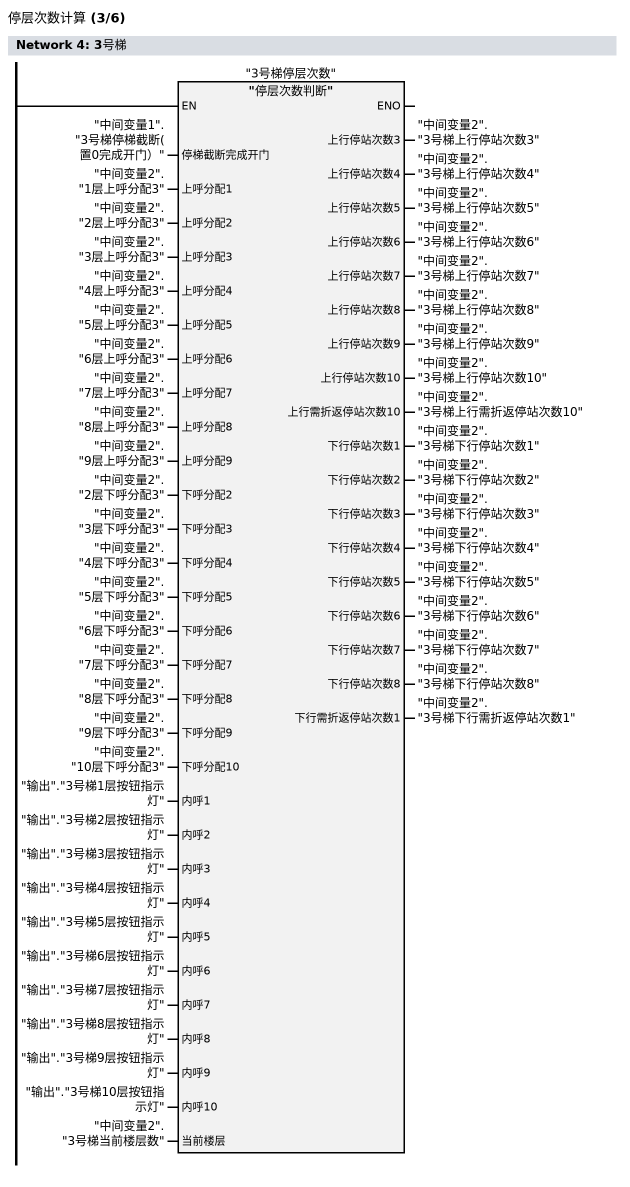
   RUNG wire#powerrail
      "3号梯停层次数"(停梯截断完成开门 := "中间变量1"."3号梯停梯截断(置0完成开门）", 上呼分配1 := "中间变量2"."1层上呼分配3", 上呼分配2 := "中间变量2"."2层上呼分配3", 上呼分配3 := "中间变量2"."3层上呼分配3", 上呼分配4 := "中间变量2"."4层上呼分配3", 上呼分配5 := "中间变量2"."5层上呼分配3", 上呼分配6 := "中间变量2"."6层上呼分配3", 上呼分配7 := "中间变量2"."7层上呼分配3", 上呼分配8 := "中间变量2"."8层上呼分配3", 上呼分配9 := "中间变量2"."9层上呼分配3", 下呼分配2 := "中间变量2"."2层下呼分配3", 下呼分配3 := "中间变量2"."3层下呼分配3", 下呼分配4 := "中间变量2"."4层下呼分配3", 下呼分配5 := "中间变量2"."5层下呼分配3", 下呼分配6 := "中间变量2"."6层下呼分配3", 下呼分配7 := "中间变量2"."7层下呼分配3", 下呼分配8 := "中间变量2"."8层下呼分配3", 下呼分配9 := "中间变量2"."9层下呼分配3", 下呼分配10 := "中间变量2"."10层下呼分配3", 内呼1 := "输出"."3号梯1层按钮指示灯", 内呼2 := "输出"."3号梯2层按钮指示灯", 内呼3 := "输出"."3号梯3层按钮指示灯", 内呼4 := "输出"."3号梯4层按钮指示灯", 内呼5 := "输出"."3号梯5层按钮指示灯", 内呼6 := "输出"."3号梯6层按钮指示灯", 内呼7 := "输出"."3号梯7层按钮指示灯", 内呼8 := "输出"."3号梯8层按钮指示灯", 内呼9 := "输出"."3号梯9层按钮指示灯", 内呼10 := "输出"."3号梯10层按钮指示灯", 当前楼层 := "中间变量2"."3号梯当前楼层数", 上行停站次数3 => "中间变量2"."3号梯上行停站次数3", 上行停站次数4 => "中间变量2"."3号梯上行停站次数4", 上行停站次数5 => "中间变量2"."3号梯上行停站次数5", 上行停站次数6 => "中间变量2"."3号梯上行停站次数6", 上行停站次数7 => "中间变量2"."3号梯上行停站次数7", 上行停站次数8 => "中间变量2"."3号梯上行停站次数8", 上行停站次数9 => "中间变量2"."3号梯上行停站次数9", 上行停站次数10 => "中间变量2"."3号梯上行停站次数10", 上行需折返停站次数10 => "中间变量2"."3号梯上行需折返停站次数10", 下行停站次数1 => "中间变量2"."3号梯下行停站次数1", 下行停站次数2 => "中间变量2"."3号梯下行停站次数2", 下行停站次数3 => "中间变量2"."3号梯下行停站次数3", 下行停站次数4 => "中间变量2"."3号梯下行停站次数4", 下行停站次数5 => "中间变量2"."3号梯下行停站次数5", 下行停站次数6 => "中间变量2"."3号梯下行停站次数6", 下行停站次数7 => "中间变量2"."3号梯下行停站次数7", 下行停站次数8 => "中间变量2"."3号梯下行停站次数8", 下行需折返停站次数1 => "中间变量2"."3号梯下行需折返停站次数1")
   END_RUNG
   // the same network as SCL:
   "3号梯停层次数"(停梯截断完成开门 := "中间变量1"."3号梯停梯截断(置0完成开门）",   // "停层次数判断"
             上呼分配1 := "中间变量2"."1层上呼分配3",
             上呼分配2 := "中间变量2"."2层上呼分配3",
             上呼分配3 := "中间变量2"."3层上呼分配3",
             上呼分配4 := "中间变量2"."4层上呼分配3",
             上呼分配5 := "中间变量2"."5层上呼分配3",
             上呼分配6 := "中间变量2"."6层上呼分配3",
             上呼分配7 := "中间变量2"."7层上呼分配3",
             上呼分配8 := "中间变量2"."8层上呼分配3",
             上呼分配9 := "中间变量2"."9层上呼分配3",
             下呼分配2 := "中间变量2"."2层下呼分配3",
             下呼分配3 := "中间变量2"."3层下呼分配3",
             下呼分配4 := "中间变量2"."4层下呼分配3",
             下呼分配5 := "中间变量2"."5层下呼分配3",
             下呼分配6 := "中间变量2"."6层下呼分配3",
             下呼分配7 := "中间变量2"."7层下呼分配3",
             下呼分配8 := "中间变量2"."8层下呼分配3",
             下呼分配9 := "中间变量2"."9层下呼分配3",
             下呼分配10 := "中间变量2"."10层下呼分配3",
             内呼1 := "输出"."3号梯1层按钮指示灯",
             内呼2 := "输出"."3号梯2层按钮指示灯",
             内呼3 := "输出"."3号梯3层按钮指示灯",
             内呼4 := "输出"."3号梯4层按钮指示灯",
             内呼5 := "输出"."3号梯5层按钮指示灯",
             内呼6 := "输出"."3号梯6层按钮指示灯",
             内呼7 := "输出"."3号梯7层按钮指示灯",
             内呼8 := "输出"."3号梯8层按钮指示灯",
             内呼9 := "输出"."3号梯9层按钮指示灯",
             内呼10 := "输出"."3号梯10层按钮指示灯",
             当前楼层 := "中间变量2"."3号梯当前楼层数",
             上行停站次数3 => "中间变量2"."3号梯上行停站次数3",
             上行停站次数4 => "中间变量2"."3号梯上行停站次数4",
             上行停站次数5 => "中间变量2"."3号梯上行停站次数5",
             上行停站次数6 => "中间变量2"."3号梯上行停站次数6",
             上行停站次数7 => "中间变量2"."3号梯上行停站次数7",
             上行停站次数8 => "中间变量2"."3号梯上行停站次数8",
             上行停站次数9 => "中间变量2"."3号梯上行停站次数9",
             上行停站次数10 => "中间变量2"."3号梯上行停站次数10",
             上行需折返停站次数10 => "中间变量2"."3号梯上行需折返停站次数10",
             下行停站次数1 => "中间变量2"."3号梯下行停站次数1",
             下行停站次数2 => "中间变量2"."3号梯下行停站次数2",
             下行停站次数3 => "中间变量2"."3号梯下行停站次数3",
             下行停站次数4 => "中间变量2"."3号梯下行停站次数4",
             下行停站次数5 => "中间变量2"."3号梯下行停站次数5",
             下行停站次数6 => "中间变量2"."3号梯下行停站次数6",
             下行停站次数7 => "中间变量2"."3号梯下行停站次数7",
             下行停站次数8 => "中间变量2"."3号梯下行停站次数8",
             下行需折返停站次数1 => "中间变量2"."3号梯下行需折返停站次数1");
END_REGION

REGION Network 5: 4号梯
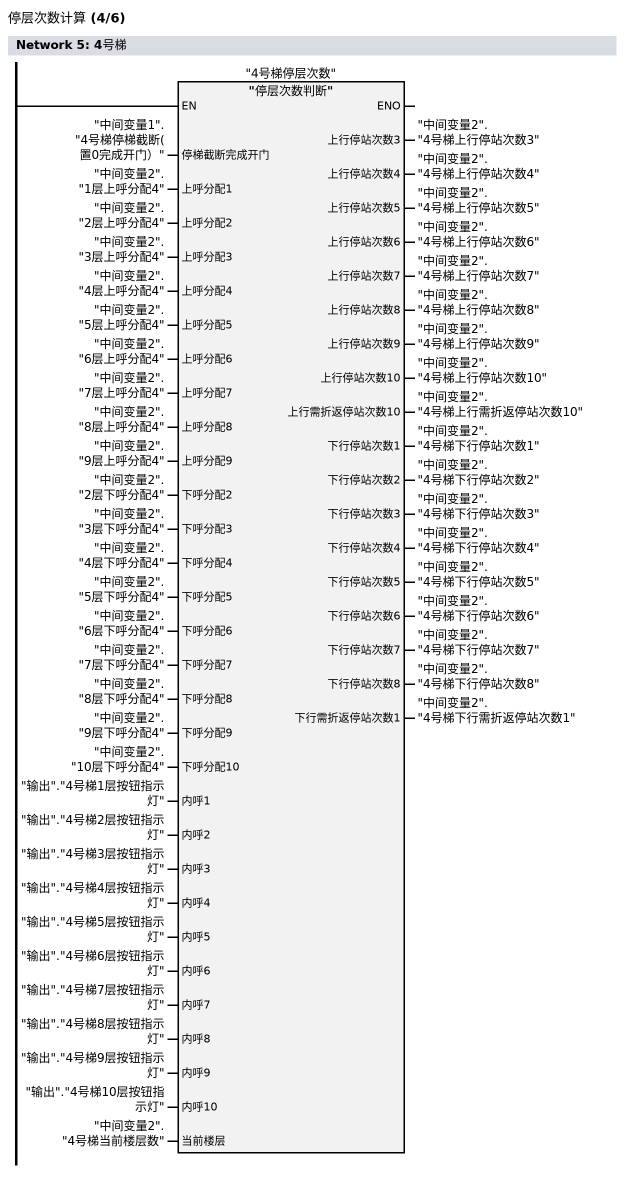
   RUNG wire#powerrail
      "4号梯停层次数"(停梯截断完成开门 := "中间变量1"."4号梯停梯截断(置0完成开门）", 上呼分配1 := "中间变量2"."1层上呼分配4", 上呼分配2 := "中间变量2"."2层上呼分配4", 上呼分配3 := "中间变量2"."3层上呼分配4", 上呼分配4 := "中间变量2"."4层上呼分配4", 上呼分配5 := "中间变量2"."5层上呼分配4", 上呼分配6 := "中间变量2"."6层上呼分配4", 上呼分配7 := "中间变量2"."7层上呼分配4", 上呼分配8 := "中间变量2"."8层上呼分配4", 上呼分配9 := "中间变量2"."9层上呼分配4", 下呼分配2 := "中间变量2"."2层下呼分配4", 下呼分配3 := "中间变量2"."3层下呼分配4", 下呼分配4 := "中间变量2"."4层下呼分配4", 下呼分配5 := "中间变量2"."5层下呼分配4", 下呼分配6 := "中间变量2"."6层下呼分配4", 下呼分配7 := "中间变量2"."7层下呼分配4", 下呼分配8 := "中间变量2"."8层下呼分配4", 下呼分配9 := "中间变量2"."9层下呼分配4", 下呼分配10 := "中间变量2"."10层下呼分配4", 内呼1 := "输出"."4号梯1层按钮指示灯", 内呼2 := "输出"."4号梯2层按钮指示灯", 内呼3 := "输出"."4号梯3层按钮指示灯", 内呼4 := "输出"."4号梯4层按钮指示灯", 内呼5 := "输出"."4号梯5层按钮指示灯", 内呼6 := "输出"."4号梯6层按钮指示灯", 内呼7 := "输出"."4号梯7层按钮指示灯", 内呼8 := "输出"."4号梯8层按钮指示灯", 内呼9 := "输出"."4号梯9层按钮指示灯", 内呼10 := "输出"."4号梯10层按钮指示灯", 当前楼层 := "中间变量2"."4号梯当前楼层数", 上行停站次数3 => "中间变量2"."4号梯上行停站次数3", 上行停站次数4 => "中间变量2"."4号梯上行停站次数4", 上行停站次数5 => "中间变量2"."4号梯上行停站次数5", 上行停站次数6 => "中间变量2"."4号梯上行停站次数6", 上行停站次数7 => "中间变量2"."4号梯上行停站次数7", 上行停站次数8 => "中间变量2"."4号梯上行停站次数8", 上行停站次数9 => "中间变量2"."4号梯上行停站次数9", 上行停站次数10 => "中间变量2"."4号梯上行停站次数10", 上行需折返停站次数10 => "中间变量2"."4号梯上行需折返停站次数10", 下行停站次数1 => "中间变量2"."4号梯下行停站次数1", 下行停站次数2 => "中间变量2"."4号梯下行停站次数2", 下行停站次数3 => "中间变量2"."4号梯下行停站次数3", 下行停站次数4 => "中间变量2"."4号梯下行停站次数4", 下行停站次数5 => "中间变量2"."4号梯下行停站次数5", 下行停站次数6 => "中间变量2"."4号梯下行停站次数6", 下行停站次数7 => "中间变量2"."4号梯下行停站次数7", 下行停站次数8 => "中间变量2"."4号梯下行停站次数8", 下行需折返停站次数1 => "中间变量2"."4号梯下行需折返停站次数1")
   END_RUNG
   // the same network as SCL:
   "4号梯停层次数"(停梯截断完成开门 := "中间变量1"."4号梯停梯截断(置0完成开门）",   // "停层次数判断"
             上呼分配1 := "中间变量2"."1层上呼分配4",
             上呼分配2 := "中间变量2"."2层上呼分配4",
             上呼分配3 := "中间变量2"."3层上呼分配4",
             上呼分配4 := "中间变量2"."4层上呼分配4",
             上呼分配5 := "中间变量2"."5层上呼分配4",
             上呼分配6 := "中间变量2"."6层上呼分配4",
             上呼分配7 := "中间变量2"."7层上呼分配4",
             上呼分配8 := "中间变量2"."8层上呼分配4",
             上呼分配9 := "中间变量2"."9层上呼分配4",
             下呼分配2 := "中间变量2"."2层下呼分配4",
             下呼分配3 := "中间变量2"."3层下呼分配4",
             下呼分配4 := "中间变量2"."4层下呼分配4",
             下呼分配5 := "中间变量2"."5层下呼分配4",
             下呼分配6 := "中间变量2"."6层下呼分配4",
             下呼分配7 := "中间变量2"."7层下呼分配4",
             下呼分配8 := "中间变量2"."8层下呼分配4",
             下呼分配9 := "中间变量2"."9层下呼分配4",
             下呼分配10 := "中间变量2"."10层下呼分配4",
             内呼1 := "输出"."4号梯1层按钮指示灯",
             内呼2 := "输出"."4号梯2层按钮指示灯",
             内呼3 := "输出"."4号梯3层按钮指示灯",
             内呼4 := "输出"."4号梯4层按钮指示灯",
             内呼5 := "输出"."4号梯5层按钮指示灯",
             内呼6 := "输出"."4号梯6层按钮指示灯",
             内呼7 := "输出"."4号梯7层按钮指示灯",
             内呼8 := "输出"."4号梯8层按钮指示灯",
             内呼9 := "输出"."4号梯9层按钮指示灯",
             内呼10 := "输出"."4号梯10层按钮指示灯",
             当前楼层 := "中间变量2"."4号梯当前楼层数",
             上行停站次数3 => "中间变量2"."4号梯上行停站次数3",
             上行停站次数4 => "中间变量2"."4号梯上行停站次数4",
             上行停站次数5 => "中间变量2"."4号梯上行停站次数5",
             上行停站次数6 => "中间变量2"."4号梯上行停站次数6",
             上行停站次数7 => "中间变量2"."4号梯上行停站次数7",
             上行停站次数8 => "中间变量2"."4号梯上行停站次数8",
             上行停站次数9 => "中间变量2"."4号梯上行停站次数9",
             上行停站次数10 => "中间变量2"."4号梯上行停站次数10",
             上行需折返停站次数10 => "中间变量2"."4号梯上行需折返停站次数10",
             下行停站次数1 => "中间变量2"."4号梯下行停站次数1",
             下行停站次数2 => "中间变量2"."4号梯下行停站次数2",
             下行停站次数3 => "中间变量2"."4号梯下行停站次数3",
             下行停站次数4 => "中间变量2"."4号梯下行停站次数4",
             下行停站次数5 => "中间变量2"."4号梯下行停站次数5",
             下行停站次数6 => "中间变量2"."4号梯下行停站次数6",
             下行停站次数7 => "中间变量2"."4号梯下行停站次数7",
             下行停站次数8 => "中间变量2"."4号梯下行停站次数8",
             下行需折返停站次数1 => "中间变量2"."4号梯下行需折返停站次数1");
END_REGION

REGION Network 6: 5号梯
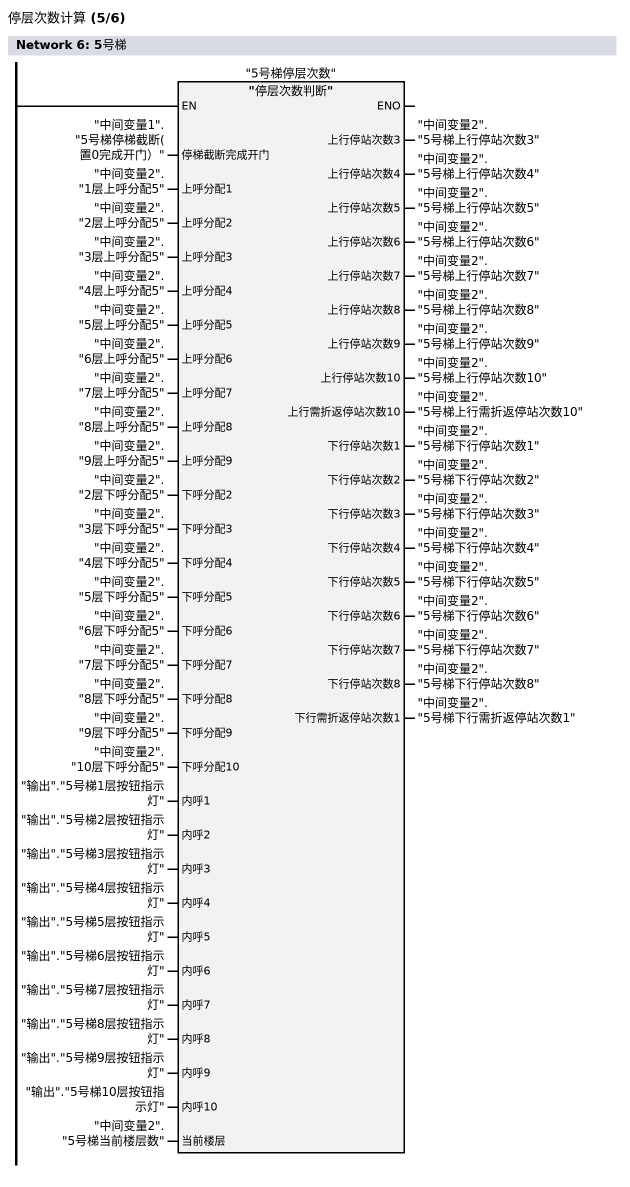
   RUNG wire#powerrail
      "5号梯停层次数"(停梯截断完成开门 := "中间变量1"."5号梯停梯截断(置0完成开门）", 上呼分配1 := "中间变量2"."1层上呼分配5", 上呼分配2 := "中间变量2"."2层上呼分配5", 上呼分配3 := "中间变量2"."3层上呼分配5", 上呼分配4 := "中间变量2"."4层上呼分配5", 上呼分配5 := "中间变量2"."5层上呼分配5", 上呼分配6 := "中间变量2"."6层上呼分配5", 上呼分配7 := "中间变量2"."7层上呼分配5", 上呼分配8 := "中间变量2"."8层上呼分配5", 上呼分配9 := "中间变量2"."9层上呼分配5", 下呼分配2 := "中间变量2"."2层下呼分配5", 下呼分配3 := "中间变量2"."3层下呼分配5", 下呼分配4 := "中间变量2"."4层下呼分配5", 下呼分配5 := "中间变量2"."5层下呼分配5", 下呼分配6 := "中间变量2"."6层下呼分配5", 下呼分配7 := "中间变量2"."7层下呼分配5", 下呼分配8 := "中间变量2"."8层下呼分配5", 下呼分配9 := "中间变量2"."9层下呼分配5", 下呼分配10 := "中间变量2"."10层下呼分配5", 内呼1 := "输出"."5号梯1层按钮指示灯", 内呼2 := "输出"."5号梯2层按钮指示灯", 内呼3 := "输出"."5号梯3层按钮指示灯", 内呼4 := "输出"."5号梯4层按钮指示灯", 内呼5 := "输出"."5号梯5层按钮指示灯", 内呼6 := "输出"."5号梯6层按钮指示灯", 内呼7 := "输出"."5号梯7层按钮指示灯", 内呼8 := "输出"."5号梯8层按钮指示灯", 内呼9 := "输出"."5号梯9层按钮指示灯", 内呼10 := "输出"."5号梯10层按钮指示灯", 当前楼层 := "中间变量2"."5号梯当前楼层数", 上行停站次数3 => "中间变量2"."5号梯上行停站次数3", 上行停站次数4 => "中间变量2"."5号梯上行停站次数4", 上行停站次数5 => "中间变量2"."5号梯上行停站次数5", 上行停站次数6 => "中间变量2"."5号梯上行停站次数6", 上行停站次数7 => "中间变量2"."5号梯上行停站次数7", 上行停站次数8 => "中间变量2"."5号梯上行停站次数8", 上行停站次数9 => "中间变量2"."5号梯上行停站次数9", 上行停站次数10 => "中间变量2"."5号梯上行停站次数10", 上行需折返停站次数10 => "中间变量2"."5号梯上行需折返停站次数10", 下行停站次数1 => "中间变量2"."5号梯下行停站次数1", 下行停站次数2 => "中间变量2"."5号梯下行停站次数2", 下行停站次数3 => "中间变量2"."5号梯下行停站次数3", 下行停站次数4 => "中间变量2"."5号梯下行停站次数4", 下行停站次数5 => "中间变量2"."5号梯下行停站次数5", 下行停站次数6 => "中间变量2"."5号梯下行停站次数6", 下行停站次数7 => "中间变量2"."5号梯下行停站次数7", 下行停站次数8 => "中间变量2"."5号梯下行停站次数8", 下行需折返停站次数1 => "中间变量2"."5号梯下行需折返停站次数1")
   END_RUNG
   // the same network as SCL:
   "5号梯停层次数"(停梯截断完成开门 := "中间变量1"."5号梯停梯截断(置0完成开门）",   // "停层次数判断"
             上呼分配1 := "中间变量2"."1层上呼分配5",
             上呼分配2 := "中间变量2"."2层上呼分配5",
             上呼分配3 := "中间变量2"."3层上呼分配5",
             上呼分配4 := "中间变量2"."4层上呼分配5",
             上呼分配5 := "中间变量2"."5层上呼分配5",
             上呼分配6 := "中间变量2"."6层上呼分配5",
             上呼分配7 := "中间变量2"."7层上呼分配5",
             上呼分配8 := "中间变量2"."8层上呼分配5",
             上呼分配9 := "中间变量2"."9层上呼分配5",
             下呼分配2 := "中间变量2"."2层下呼分配5",
             下呼分配3 := "中间变量2"."3层下呼分配5",
             下呼分配4 := "中间变量2"."4层下呼分配5",
             下呼分配5 := "中间变量2"."5层下呼分配5",
             下呼分配6 := "中间变量2"."6层下呼分配5",
             下呼分配7 := "中间变量2"."7层下呼分配5",
             下呼分配8 := "中间变量2"."8层下呼分配5",
             下呼分配9 := "中间变量2"."9层下呼分配5",
             下呼分配10 := "中间变量2"."10层下呼分配5",
             内呼1 := "输出"."5号梯1层按钮指示灯",
             内呼2 := "输出"."5号梯2层按钮指示灯",
             内呼3 := "输出"."5号梯3层按钮指示灯",
             内呼4 := "输出"."5号梯4层按钮指示灯",
             内呼5 := "输出"."5号梯5层按钮指示灯",
             内呼6 := "输出"."5号梯6层按钮指示灯",
             内呼7 := "输出"."5号梯7层按钮指示灯",
             内呼8 := "输出"."5号梯8层按钮指示灯",
             内呼9 := "输出"."5号梯9层按钮指示灯",
             内呼10 := "输出"."5号梯10层按钮指示灯",
             当前楼层 := "中间变量2"."5号梯当前楼层数",
             上行停站次数3 => "中间变量2"."5号梯上行停站次数3",
             上行停站次数4 => "中间变量2"."5号梯上行停站次数4",
             上行停站次数5 => "中间变量2"."5号梯上行停站次数5",
             上行停站次数6 => "中间变量2"."5号梯上行停站次数6",
             上行停站次数7 => "中间变量2"."5号梯上行停站次数7",
             上行停站次数8 => "中间变量2"."5号梯上行停站次数8",
             上行停站次数9 => "中间变量2"."5号梯上行停站次数9",
             上行停站次数10 => "中间变量2"."5号梯上行停站次数10",
             上行需折返停站次数10 => "中间变量2"."5号梯上行需折返停站次数10",
             下行停站次数1 => "中间变量2"."5号梯下行停站次数1",
             下行停站次数2 => "中间变量2"."5号梯下行停站次数2",
             下行停站次数3 => "中间变量2"."5号梯下行停站次数3",
             下行停站次数4 => "中间变量2"."5号梯下行停站次数4",
             下行停站次数5 => "中间变量2"."5号梯下行停站次数5",
             下行停站次数6 => "中间变量2"."5号梯下行停站次数6",
             下行停站次数7 => "中间变量2"."5号梯下行停站次数7",
             下行停站次数8 => "中间变量2"."5号梯下行停站次数8",
             下行需折返停站次数1 => "中间变量2"."5号梯下行需折返停站次数1");
END_REGION

REGION Network 7: 6号梯
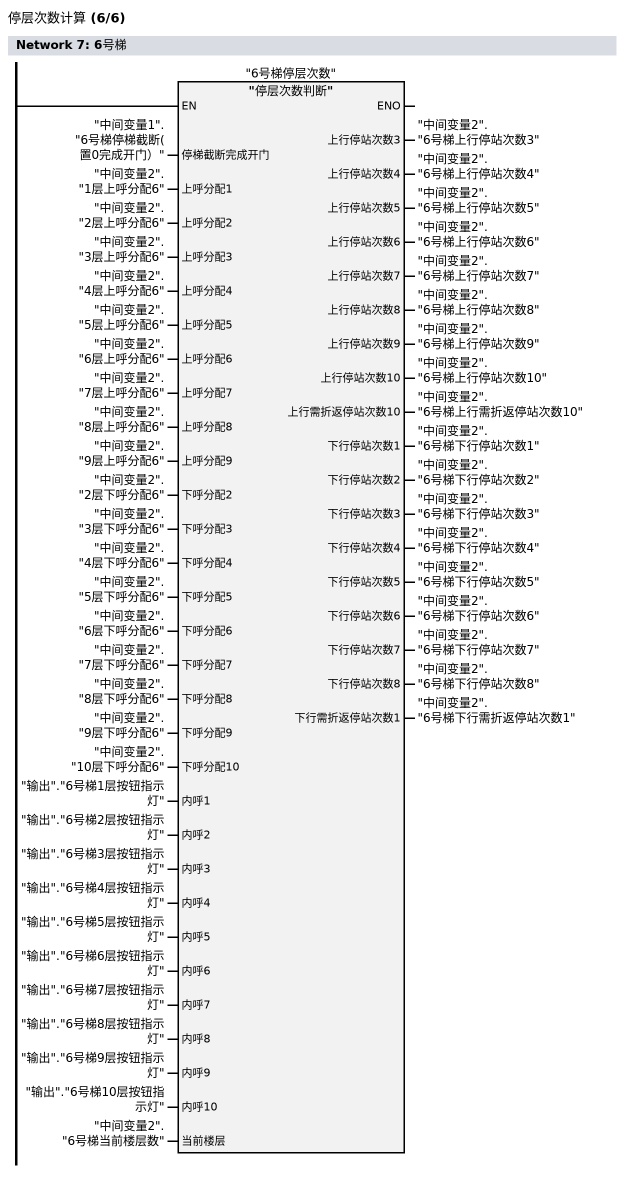
   RUNG wire#powerrail
      "6号梯停层次数"(停梯截断完成开门 := "中间变量1"."6号梯停梯截断(置0完成开门）", 上呼分配1 := "中间变量2"."1层上呼分配6", 上呼分配2 := "中间变量2"."2层上呼分配6", 上呼分配3 := "中间变量2"."3层上呼分配6", 上呼分配4 := "中间变量2"."4层上呼分配6", 上呼分配5 := "中间变量2"."5层上呼分配6", 上呼分配6 := "中间变量2"."6层上呼分配6", 上呼分配7 := "中间变量2"."7层上呼分配6", 上呼分配8 := "中间变量2"."8层上呼分配6", 上呼分配9 := "中间变量2"."9层上呼分配6", 下呼分配2 := "中间变量2"."2层下呼分配6", 下呼分配3 := "中间变量2"."3层下呼分配6", 下呼分配4 := "中间变量2"."4层下呼分配6", 下呼分配5 := "中间变量2"."5层下呼分配6", 下呼分配6 := "中间变量2"."6层下呼分配6", 下呼分配7 := "中间变量2"."7层下呼分配6", 下呼分配8 := "中间变量2"."8层下呼分配6", 下呼分配9 := "中间变量2"."9层下呼分配6", 下呼分配10 := "中间变量2"."10层下呼分配6", 内呼1 := "输出"."6号梯1层按钮指示灯", 内呼2 := "输出"."6号梯2层按钮指示灯", 内呼3 := "输出"."6号梯3层按钮指示灯", 内呼4 := "输出"."6号梯4层按钮指示灯", 内呼5 := "输出"."6号梯5层按钮指示灯", 内呼6 := "输出"."6号梯6层按钮指示灯", 内呼7 := "输出"."6号梯7层按钮指示灯", 内呼8 := "输出"."6号梯8层按钮指示灯", 内呼9 := "输出"."6号梯9层按钮指示灯", 内呼10 := "输出"."6号梯10层按钮指示灯", 当前楼层 := "中间变量2"."6号梯当前楼层数", 上行停站次数3 => "中间变量2"."6号梯上行停站次数3", 上行停站次数4 => "中间变量2"."6号梯上行停站次数4", 上行停站次数5 => "中间变量2"."6号梯上行停站次数5", 上行停站次数6 => "中间变量2"."6号梯上行停站次数6", 上行停站次数7 => "中间变量2"."6号梯上行停站次数7", 上行停站次数8 => "中间变量2"."6号梯上行停站次数8", 上行停站次数9 => "中间变量2"."6号梯上行停站次数9", 上行停站次数10 => "中间变量2"."6号梯上行停站次数10", 上行需折返停站次数10 => "中间变量2"."6号梯上行需折返停站次数10", 下行停站次数1 => "中间变量2"."6号梯下行停站次数1", 下行停站次数2 => "中间变量2"."6号梯下行停站次数2", 下行停站次数3 => "中间变量2"."6号梯下行停站次数3", 下行停站次数4 => "中间变量2"."6号梯下行停站次数4", 下行停站次数5 => "中间变量2"."6号梯下行停站次数5", 下行停站次数6 => "中间变量2"."6号梯下行停站次数6", 下行停站次数7 => "中间变量2"."6号梯下行停站次数7", 下行停站次数8 => "中间变量2"."6号梯下行停站次数8", 下行需折返停站次数1 => "中间变量2"."6号梯下行需折返停站次数1")
   END_RUNG
   // the same network as SCL:
   "6号梯停层次数"(停梯截断完成开门 := "中间变量1"."6号梯停梯截断(置0完成开门）",   // "停层次数判断"
             上呼分配1 := "中间变量2"."1层上呼分配6",
             上呼分配2 := "中间变量2"."2层上呼分配6",
             上呼分配3 := "中间变量2"."3层上呼分配6",
             上呼分配4 := "中间变量2"."4层上呼分配6",
             上呼分配5 := "中间变量2"."5层上呼分配6",
             上呼分配6 := "中间变量2"."6层上呼分配6",
             上呼分配7 := "中间变量2"."7层上呼分配6",
             上呼分配8 := "中间变量2"."8层上呼分配6",
             上呼分配9 := "中间变量2"."9层上呼分配6",
             下呼分配2 := "中间变量2"."2层下呼分配6",
             下呼分配3 := "中间变量2"."3层下呼分配6",
             下呼分配4 := "中间变量2"."4层下呼分配6",
             下呼分配5 := "中间变量2"."5层下呼分配6",
             下呼分配6 := "中间变量2"."6层下呼分配6",
             下呼分配7 := "中间变量2"."7层下呼分配6",
             下呼分配8 := "中间变量2"."8层下呼分配6",
             下呼分配9 := "中间变量2"."9层下呼分配6",
             下呼分配10 := "中间变量2"."10层下呼分配6",
             内呼1 := "输出"."6号梯1层按钮指示灯",
             内呼2 := "输出"."6号梯2层按钮指示灯",
             内呼3 := "输出"."6号梯3层按钮指示灯",
             内呼4 := "输出"."6号梯4层按钮指示灯",
             内呼5 := "输出"."6号梯5层按钮指示灯",
             内呼6 := "输出"."6号梯6层按钮指示灯",
             内呼7 := "输出"."6号梯7层按钮指示灯",
             内呼8 := "输出"."6号梯8层按钮指示灯",
             内呼9 := "输出"."6号梯9层按钮指示灯",
             内呼10 := "输出"."6号梯10层按钮指示灯",
             当前楼层 := "中间变量2"."6号梯当前楼层数",
             上行停站次数3 => "中间变量2"."6号梯上行停站次数3",
             上行停站次数4 => "中间变量2"."6号梯上行停站次数4",
             上行停站次数5 => "中间变量2"."6号梯上行停站次数5",
             上行停站次数6 => "中间变量2"."6号梯上行停站次数6",
             上行停站次数7 => "中间变量2"."6号梯上行停站次数7",
             上行停站次数8 => "中间变量2"."6号梯上行停站次数8",
             上行停站次数9 => "中间变量2"."6号梯上行停站次数9",
             上行停站次数10 => "中间变量2"."6号梯上行停站次数10",
             上行需折返停站次数10 => "中间变量2"."6号梯上行需折返停站次数10",
             下行停站次数1 => "中间变量2"."6号梯下行停站次数1",
             下行停站次数2 => "中间变量2"."6号梯下行停站次数2",
             下行停站次数3 => "中间变量2"."6号梯下行停站次数3",
             下行停站次数4 => "中间变量2"."6号梯下行停站次数4",
             下行停站次数5 => "中间变量2"."6号梯下行停站次数5",
             下行停站次数6 => "中间变量2"."6号梯下行停站次数6",
             下行停站次数7 => "中间变量2"."6号梯下行停站次数7",
             下行停站次数8 => "中间变量2"."6号梯下行停站次数8",
             下行需折返停站次数1 => "中间变量2"."6号梯下行需折返停站次数1");
END_REGION
END_FUNCTION

FUNCTION "初始化赋值" : Void   // FC8, LAD
{ S7_Optimized_Access := 'TRUE' }
VERSION : 0.1
   VAR_TEMP   // added for the SCL form of the ladder/FBD networks
      _w1 : Bool;
      _w2 : Bool;
      _w3 : Bool;
      _w4 : Bool;
      _w5 : Bool;
      _w6 : Bool;
   END_VAR
BEGIN

REGION Network 1: 初始化楼层
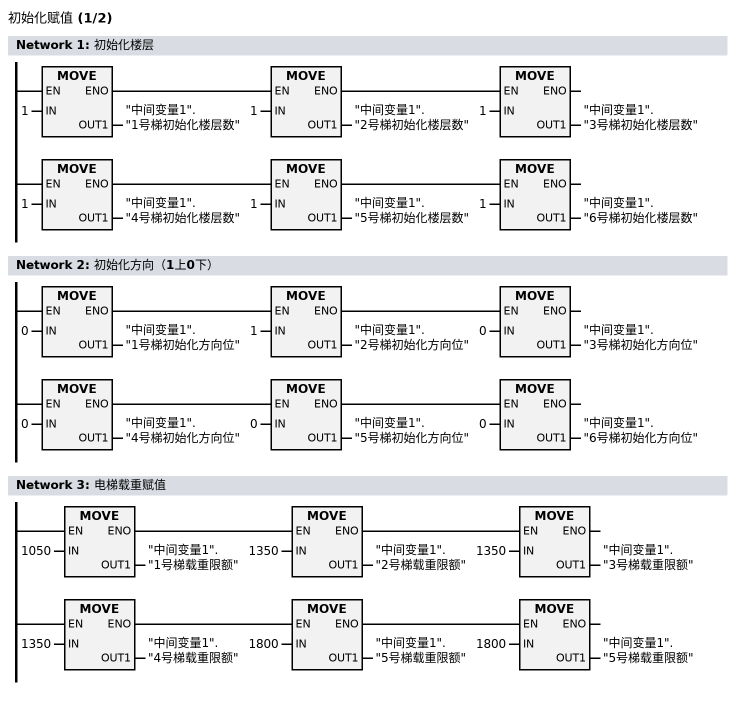
   RUNG wire#powerrail
      Move(in := 1, out1 => "中间变量1"."1号梯初始化楼层数")
      Move(in := 1, out1 => "中间变量1"."2号梯初始化楼层数")
      Move(in := 1, out1 => "中间变量1"."3号梯初始化楼层数")
   END_RUNG
   RUNG wire#powerrail
      Move(in := 1, out1 => "中间变量1"."4号梯初始化楼层数")
      Move(in := 1, out1 => "中间变量1"."5号梯初始化楼层数")
      Move(in := 1, out1 => "中间变量1"."6号梯初始化楼层数")
   END_RUNG
   // the same network as SCL:
   "中间变量1"."1号梯初始化楼层数" := 1;
   "中间变量1"."2号梯初始化楼层数" := 1;
   "中间变量1"."3号梯初始化楼层数" := 1;
   "中间变量1"."4号梯初始化楼层数" := 1;
   "中间变量1"."5号梯初始化楼层数" := 1;
   "中间变量1"."6号梯初始化楼层数" := 1;
END_REGION

REGION Network 2: 初始化方向（1上0下）
   RUNG wire#powerrail
      Move(in := 0, out1 => "中间变量1"."1号梯初始化方向位")
      Move(in := 1, out1 => "中间变量1"."2号梯初始化方向位")
      Move(in := 0, out1 => "中间变量1"."3号梯初始化方向位")
   END_RUNG
   RUNG wire#powerrail
      Move(in := 0, out1 => "中间变量1"."4号梯初始化方向位")
      Move(in := 0, out1 => "中间变量1"."5号梯初始化方向位")
      Move(in := 0, out1 => "中间变量1"."6号梯初始化方向位")
   END_RUNG
   // the same network as SCL:
   "中间变量1"."1号梯初始化方向位" := 0;
   "中间变量1"."2号梯初始化方向位" := 1;
   "中间变量1"."3号梯初始化方向位" := 0;
   "中间变量1"."4号梯初始化方向位" := 0;
   "中间变量1"."5号梯初始化方向位" := 0;
   "中间变量1"."6号梯初始化方向位" := 0;
END_REGION

REGION Network 3: 电梯载重赋值
   RUNG wire#powerrail
      Move(in := 1050, out1 => "中间变量1"."1号梯载重限额")
      Move(in := 1350, out1 => "中间变量1"."2号梯载重限额")
      Move(in := 1350, out1 => "中间变量1"."3号梯载重限额")
   END_RUNG
   RUNG wire#powerrail
      Move(in := 1350, out1 => "中间变量1"."4号梯载重限额")
      Move(in := 1800, out1 => "中间变量1"."5号梯载重限额")
      Move(in := 1800, out1 => "中间变量1"."5号梯载重限额")
   END_RUNG
   // the same network as SCL:
   "中间变量1"."1号梯载重限额" := 1050;
   "中间变量1"."2号梯载重限额" := 1350;
   "中间变量1"."3号梯载重限额" := 1350;
   "中间变量1"."4号梯载重限额" := 1350;
   "中间变量1"."5号梯载重限额" := 1800;
   "中间变量1"."5号梯载重限额" := 1800;
END_REGION

REGION Network 4: 初始化方向执行
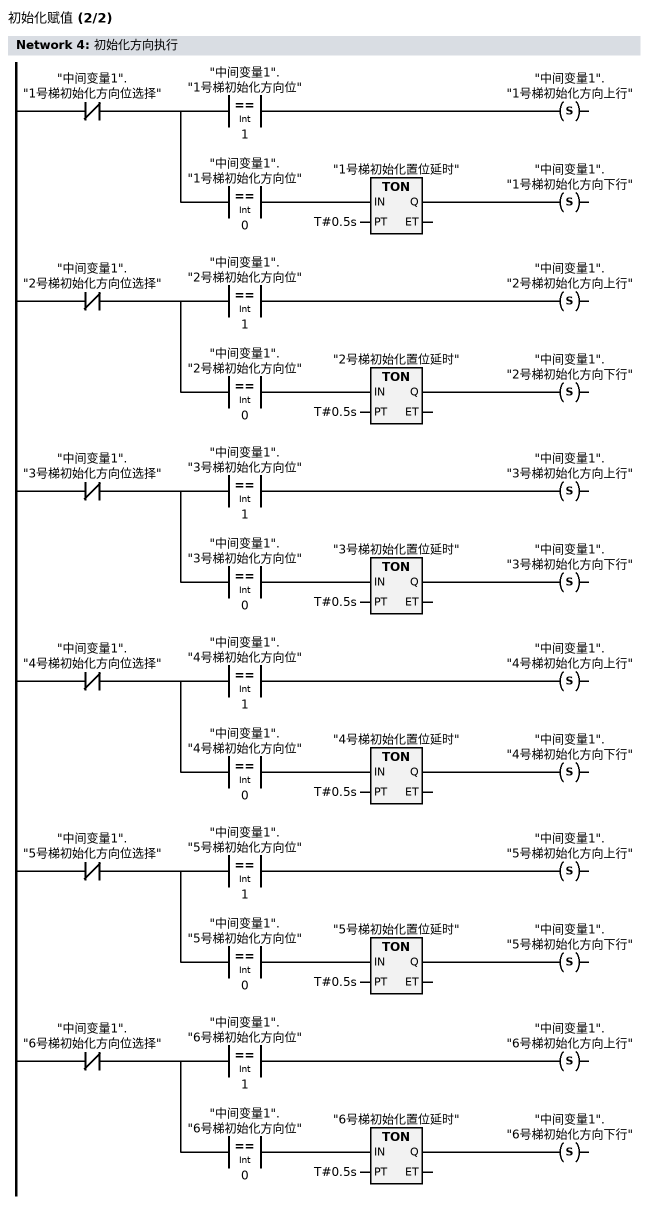
   #_w1 := NOT "中间变量1"."1号梯初始化方向位选择";
   IF #_w1 AND ("中间变量1"."1号梯初始化方向位" = 1) THEN "中间变量1"."1号梯初始化方向上行" := TRUE; END_IF;
   "1号梯初始化置位延时".TON(IN := #_w1 AND ("中间变量1"."1号梯初始化方向位" = 0), PT := T#0.5s);
   IF "1号梯初始化置位延时".Q THEN "中间变量1"."1号梯初始化方向下行" := TRUE; END_IF;
   #_w2 := NOT "中间变量1"."2号梯初始化方向位选择";
   IF #_w2 AND ("中间变量1"."2号梯初始化方向位" = 1) THEN "中间变量1"."2号梯初始化方向上行" := TRUE; END_IF;
   "2号梯初始化置位延时".TON(IN := #_w2 AND ("中间变量1"."2号梯初始化方向位" = 0), PT := T#0.5s);
   IF "2号梯初始化置位延时".Q THEN "中间变量1"."2号梯初始化方向下行" := TRUE; END_IF;
   #_w3 := NOT "中间变量1"."3号梯初始化方向位选择";
   IF #_w3 AND ("中间变量1"."3号梯初始化方向位" = 1) THEN "中间变量1"."3号梯初始化方向上行" := TRUE; END_IF;
   "3号梯初始化置位延时".TON(IN := #_w3 AND ("中间变量1"."3号梯初始化方向位" = 0), PT := T#0.5s);
   IF "3号梯初始化置位延时".Q THEN "中间变量1"."3号梯初始化方向下行" := TRUE; END_IF;
   #_w4 := NOT "中间变量1"."4号梯初始化方向位选择";
   IF #_w4 AND ("中间变量1"."4号梯初始化方向位" = 1) THEN "中间变量1"."4号梯初始化方向上行" := TRUE; END_IF;
   "4号梯初始化置位延时".TON(IN := #_w4 AND ("中间变量1"."4号梯初始化方向位" = 0), PT := T#0.5s);
   IF "4号梯初始化置位延时".Q THEN "中间变量1"."4号梯初始化方向下行" := TRUE; END_IF;
   #_w5 := NOT "中间变量1"."5号梯初始化方向位选择";
   IF #_w5 AND ("中间变量1"."5号梯初始化方向位" = 1) THEN "中间变量1"."5号梯初始化方向上行" := TRUE; END_IF;
   "5号梯初始化置位延时".TON(IN := #_w5 AND ("中间变量1"."5号梯初始化方向位" = 0), PT := T#0.5s);
   IF "5号梯初始化置位延时".Q THEN "中间变量1"."5号梯初始化方向下行" := TRUE; END_IF;
   #_w6 := NOT "中间变量1"."6号梯初始化方向位选择";
   IF #_w6 AND ("中间变量1"."6号梯初始化方向位" = 1) THEN "中间变量1"."6号梯初始化方向上行" := TRUE; END_IF;
   "6号梯初始化置位延时".TON(IN := #_w6 AND ("中间变量1"."6号梯初始化方向位" = 0), PT := T#0.5s);
   IF "6号梯初始化置位延时".Q THEN "中间变量1"."6号梯初始化方向下行" := TRUE; END_IF;
END_REGION
END_FUNCTION

FUNCTION "楼层计数" : Void   // FC9, LAD
{ S7_Optimized_Access := 'TRUE' }
VERSION : 0.1
BEGIN

REGION Network 2
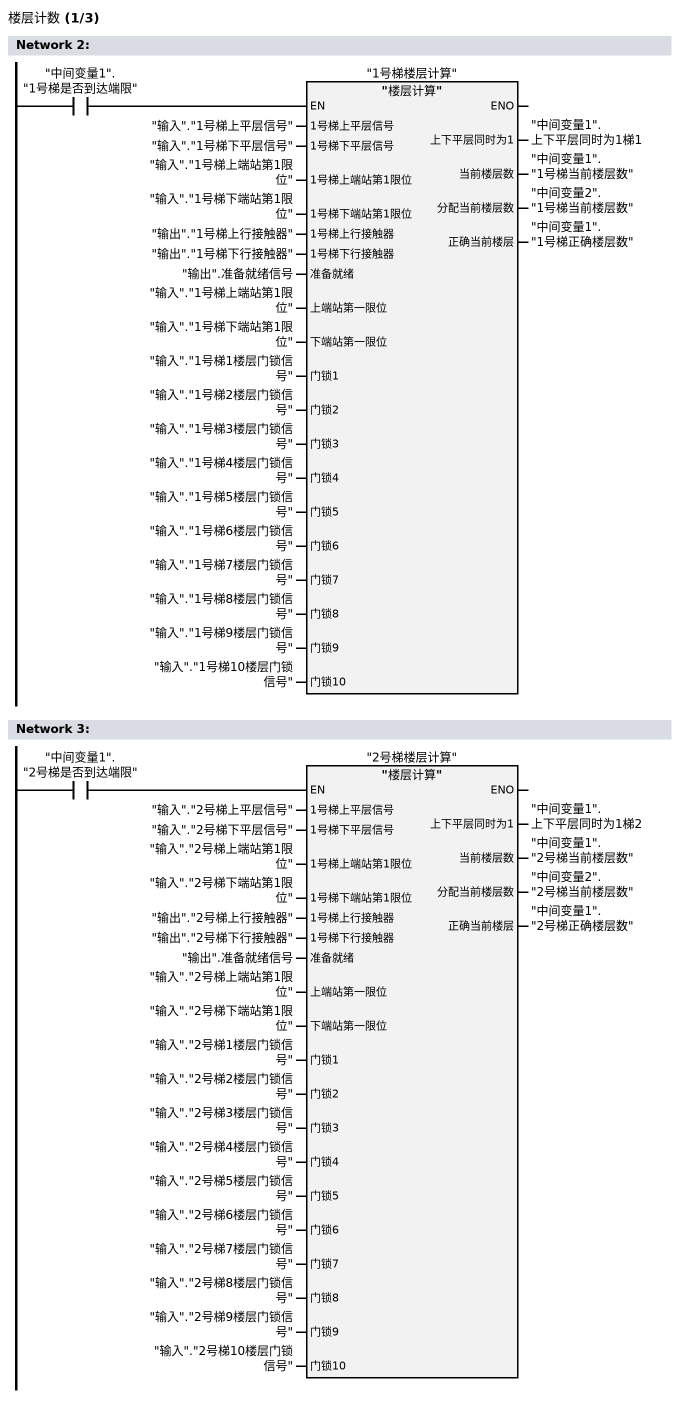
   RUNG wire#powerrail
      Contact( "中间变量1"."1号梯是否到达端限" )
      "1号梯楼层计算"("1号梯上平层信号" := "输入"."1号梯上平层信号", "1号梯下平层信号" := "输入"."1号梯下平层信号", "1号梯上端站第1限位" := "输入"."1号梯上端站第1限位", "1号梯下端站第1限位" := "输入"."1号梯下端站第1限位", "1号梯上行接触器" := "输出"."1号梯上行接触器", "1号梯下行接触器" := "输出"."1号梯下行接触器", 准备就绪 := "输出".准备就绪信号, 上端站第一限位 := "输入"."1号梯上端站第1限位", 下端站第一限位 := "输入"."1号梯下端站第1限位", 门锁1 := "输入"."1号梯1楼层门锁信号", 门锁2 := "输入"."1号梯2楼层门锁信号", 门锁3 := "输入"."1号梯3楼层门锁信号", 门锁4 := "输入"."1号梯4楼层门锁信号", 门锁5 := "输入"."1号梯5楼层门锁信号", 门锁6 := "输入"."1号梯6楼层门锁信号", 门锁7 := "输入"."1号梯7楼层门锁信号", 门锁8 := "输入"."1号梯8楼层门锁信号", 门锁9 := "输入"."1号梯9楼层门锁信号", 门锁10 := "输入"."1号梯10楼层门锁信号", 上下平层同时为1 => "中间变量1".上下平层同时为1梯1, 当前楼层数 => "中间变量1"."1号梯当前楼层数", 分配当前楼层数 => "中间变量2"."1号梯当前楼层数", 正确当前楼层 => "中间变量1"."1号梯正确楼层数")
   END_RUNG
   // the same network as SCL:
   IF "中间变量1"."1号梯是否到达端限" THEN
       "1号梯楼层计算"("1号梯上平层信号" := "输入"."1号梯上平层信号",   // "楼层计算"
                 "1号梯下平层信号" := "输入"."1号梯下平层信号",
                 "1号梯上端站第1限位" := "输入"."1号梯上端站第1限位",
                 "1号梯下端站第1限位" := "输入"."1号梯下端站第1限位",
                 "1号梯上行接触器" := "输出"."1号梯上行接触器",
                 "1号梯下行接触器" := "输出"."1号梯下行接触器",
                 准备就绪 := "输出".准备就绪信号,
                 上端站第一限位 := "输入"."1号梯上端站第1限位",
                 下端站第一限位 := "输入"."1号梯下端站第1限位",
                 门锁1 := "输入"."1号梯1楼层门锁信号",
                 门锁2 := "输入"."1号梯2楼层门锁信号",
                 门锁3 := "输入"."1号梯3楼层门锁信号",
                 门锁4 := "输入"."1号梯4楼层门锁信号",
                 门锁5 := "输入"."1号梯5楼层门锁信号",
                 门锁6 := "输入"."1号梯6楼层门锁信号",
                 门锁7 := "输入"."1号梯7楼层门锁信号",
                 门锁8 := "输入"."1号梯8楼层门锁信号",
                 门锁9 := "输入"."1号梯9楼层门锁信号",
                 门锁10 := "输入"."1号梯10楼层门锁信号",
                 上下平层同时为1 => "中间变量1".上下平层同时为1梯1,
                 当前楼层数 => "中间变量1"."1号梯当前楼层数",
                 分配当前楼层数 => "中间变量2"."1号梯当前楼层数",
                 正确当前楼层 => "中间变量1"."1号梯正确楼层数");
   END_IF;
END_REGION

REGION Network 3
   RUNG wire#powerrail
      Contact( "中间变量1"."2号梯是否到达端限" )
      "2号梯楼层计算"("1号梯上平层信号" := "输入"."2号梯上平层信号", "1号梯下平层信号" := "输入"."2号梯下平层信号", "1号梯上端站第1限位" := "输入"."2号梯上端站第1限位", "1号梯下端站第1限位" := "输入"."2号梯下端站第1限位", "1号梯上行接触器" := "输出"."2号梯上行接触器", "1号梯下行接触器" := "输出"."2号梯下行接触器", 准备就绪 := "输出".准备就绪信号, 上端站第一限位 := "输入"."2号梯上端站第1限位", 下端站第一限位 := "输入"."2号梯下端站第1限位", 门锁1 := "输入"."2号梯1楼层门锁信号", 门锁2 := "输入"."2号梯2楼层门锁信号", 门锁3 := "输入"."2号梯3楼层门锁信号", 门锁4 := "输入"."2号梯4楼层门锁信号", 门锁5 := "输入"."2号梯5楼层门锁信号", 门锁6 := "输入"."2号梯6楼层门锁信号", 门锁7 := "输入"."2号梯7楼层门锁信号", 门锁8 := "输入"."2号梯8楼层门锁信号", 门锁9 := "输入"."2号梯9楼层门锁信号", 门锁10 := "输入"."2号梯10楼层门锁信号", 上下平层同时为1 => "中间变量1".上下平层同时为1梯2, 当前楼层数 => "中间变量1"."2号梯当前楼层数", 分配当前楼层数 => "中间变量2"."2号梯当前楼层数", 正确当前楼层 => "中间变量1"."2号梯正确楼层数")
   END_RUNG
   // the same network as SCL:
   IF "中间变量1"."2号梯是否到达端限" THEN
       "2号梯楼层计算"("1号梯上平层信号" := "输入"."2号梯上平层信号",   // "楼层计算"
                 "1号梯下平层信号" := "输入"."2号梯下平层信号",
                 "1号梯上端站第1限位" := "输入"."2号梯上端站第1限位",
                 "1号梯下端站第1限位" := "输入"."2号梯下端站第1限位",
                 "1号梯上行接触器" := "输出"."2号梯上行接触器",
                 "1号梯下行接触器" := "输出"."2号梯下行接触器",
                 准备就绪 := "输出".准备就绪信号,
                 上端站第一限位 := "输入"."2号梯上端站第1限位",
                 下端站第一限位 := "输入"."2号梯下端站第1限位",
                 门锁1 := "输入"."2号梯1楼层门锁信号",
                 门锁2 := "输入"."2号梯2楼层门锁信号",
                 门锁3 := "输入"."2号梯3楼层门锁信号",
                 门锁4 := "输入"."2号梯4楼层门锁信号",
                 门锁5 := "输入"."2号梯5楼层门锁信号",
                 门锁6 := "输入"."2号梯6楼层门锁信号",
                 门锁7 := "输入"."2号梯7楼层门锁信号",
                 门锁8 := "输入"."2号梯8楼层门锁信号",
                 门锁9 := "输入"."2号梯9楼层门锁信号",
                 门锁10 := "输入"."2号梯10楼层门锁信号",
                 上下平层同时为1 => "中间变量1".上下平层同时为1梯2,
                 当前楼层数 => "中间变量1"."2号梯当前楼层数",
                 分配当前楼层数 => "中间变量2"."2号梯当前楼层数",
                 正确当前楼层 => "中间变量1"."2号梯正确楼层数");
   END_IF;
END_REGION

REGION Network 4
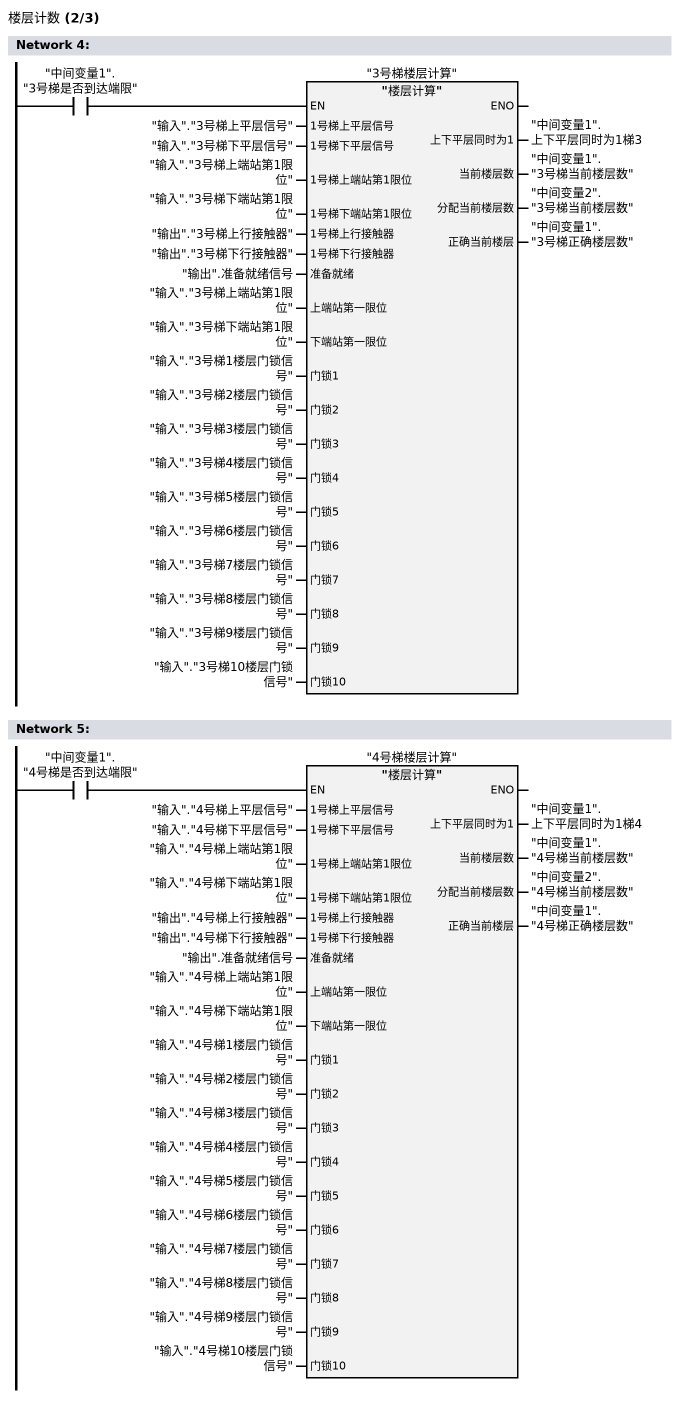
   RUNG wire#powerrail
      Contact( "中间变量1"."3号梯是否到达端限" )
      "3号梯楼层计算"("1号梯上平层信号" := "输入"."3号梯上平层信号", "1号梯下平层信号" := "输入"."3号梯下平层信号", "1号梯上端站第1限位" := "输入"."3号梯上端站第1限位", "1号梯下端站第1限位" := "输入"."3号梯下端站第1限位", "1号梯上行接触器" := "输出"."3号梯上行接触器", "1号梯下行接触器" := "输出"."3号梯下行接触器", 准备就绪 := "输出".准备就绪信号, 上端站第一限位 := "输入"."3号梯上端站第1限位", 下端站第一限位 := "输入"."3号梯下端站第1限位", 门锁1 := "输入"."3号梯1楼层门锁信号", 门锁2 := "输入"."3号梯2楼层门锁信号", 门锁3 := "输入"."3号梯3楼层门锁信号", 门锁4 := "输入"."3号梯4楼层门锁信号", 门锁5 := "输入"."3号梯5楼层门锁信号", 门锁6 := "输入"."3号梯6楼层门锁信号", 门锁7 := "输入"."3号梯7楼层门锁信号", 门锁8 := "输入"."3号梯8楼层门锁信号", 门锁9 := "输入"."3号梯9楼层门锁信号", 门锁10 := "输入"."3号梯10楼层门锁信号", 上下平层同时为1 => "中间变量1".上下平层同时为1梯3, 当前楼层数 => "中间变量1"."3号梯当前楼层数", 分配当前楼层数 => "中间变量2"."3号梯当前楼层数", 正确当前楼层 => "中间变量1"."3号梯正确楼层数")
   END_RUNG
   // the same network as SCL:
   IF "中间变量1"."3号梯是否到达端限" THEN
       "3号梯楼层计算"("1号梯上平层信号" := "输入"."3号梯上平层信号",   // "楼层计算"
                 "1号梯下平层信号" := "输入"."3号梯下平层信号",
                 "1号梯上端站第1限位" := "输入"."3号梯上端站第1限位",
                 "1号梯下端站第1限位" := "输入"."3号梯下端站第1限位",
                 "1号梯上行接触器" := "输出"."3号梯上行接触器",
                 "1号梯下行接触器" := "输出"."3号梯下行接触器",
                 准备就绪 := "输出".准备就绪信号,
                 上端站第一限位 := "输入"."3号梯上端站第1限位",
                 下端站第一限位 := "输入"."3号梯下端站第1限位",
                 门锁1 := "输入"."3号梯1楼层门锁信号",
                 门锁2 := "输入"."3号梯2楼层门锁信号",
                 门锁3 := "输入"."3号梯3楼层门锁信号",
                 门锁4 := "输入"."3号梯4楼层门锁信号",
                 门锁5 := "输入"."3号梯5楼层门锁信号",
                 门锁6 := "输入"."3号梯6楼层门锁信号",
                 门锁7 := "输入"."3号梯7楼层门锁信号",
                 门锁8 := "输入"."3号梯8楼层门锁信号",
                 门锁9 := "输入"."3号梯9楼层门锁信号",
                 门锁10 := "输入"."3号梯10楼层门锁信号",
                 上下平层同时为1 => "中间变量1".上下平层同时为1梯3,
                 当前楼层数 => "中间变量1"."3号梯当前楼层数",
                 分配当前楼层数 => "中间变量2"."3号梯当前楼层数",
                 正确当前楼层 => "中间变量1"."3号梯正确楼层数");
   END_IF;
END_REGION

REGION Network 5
   RUNG wire#powerrail
      Contact( "中间变量1"."4号梯是否到达端限" )
      "4号梯楼层计算"("1号梯上平层信号" := "输入"."4号梯上平层信号", "1号梯下平层信号" := "输入"."4号梯下平层信号", "1号梯上端站第1限位" := "输入"."4号梯上端站第1限位", "1号梯下端站第1限位" := "输入"."4号梯下端站第1限位", "1号梯上行接触器" := "输出"."4号梯上行接触器", "1号梯下行接触器" := "输出"."4号梯下行接触器", 准备就绪 := "输出".准备就绪信号, 上端站第一限位 := "输入"."4号梯上端站第1限位", 下端站第一限位 := "输入"."4号梯下端站第1限位", 门锁1 := "输入"."4号梯1楼层门锁信号", 门锁2 := "输入"."4号梯2楼层门锁信号", 门锁3 := "输入"."4号梯3楼层门锁信号", 门锁4 := "输入"."4号梯4楼层门锁信号", 门锁5 := "输入"."4号梯5楼层门锁信号", 门锁6 := "输入"."4号梯6楼层门锁信号", 门锁7 := "输入"."4号梯7楼层门锁信号", 门锁8 := "输入"."4号梯8楼层门锁信号", 门锁9 := "输入"."4号梯9楼层门锁信号", 门锁10 := "输入"."4号梯10楼层门锁信号", 上下平层同时为1 => "中间变量1".上下平层同时为1梯4, 当前楼层数 => "中间变量1"."4号梯当前楼层数", 分配当前楼层数 => "中间变量2"."4号梯当前楼层数", 正确当前楼层 => "中间变量1"."4号梯正确楼层数")
   END_RUNG
   // the same network as SCL:
   IF "中间变量1"."4号梯是否到达端限" THEN
       "4号梯楼层计算"("1号梯上平层信号" := "输入"."4号梯上平层信号",   // "楼层计算"
                 "1号梯下平层信号" := "输入"."4号梯下平层信号",
                 "1号梯上端站第1限位" := "输入"."4号梯上端站第1限位",
                 "1号梯下端站第1限位" := "输入"."4号梯下端站第1限位",
                 "1号梯上行接触器" := "输出"."4号梯上行接触器",
                 "1号梯下行接触器" := "输出"."4号梯下行接触器",
                 准备就绪 := "输出".准备就绪信号,
                 上端站第一限位 := "输入"."4号梯上端站第1限位",
                 下端站第一限位 := "输入"."4号梯下端站第1限位",
                 门锁1 := "输入"."4号梯1楼层门锁信号",
                 门锁2 := "输入"."4号梯2楼层门锁信号",
                 门锁3 := "输入"."4号梯3楼层门锁信号",
                 门锁4 := "输入"."4号梯4楼层门锁信号",
                 门锁5 := "输入"."4号梯5楼层门锁信号",
                 门锁6 := "输入"."4号梯6楼层门锁信号",
                 门锁7 := "输入"."4号梯7楼层门锁信号",
                 门锁8 := "输入"."4号梯8楼层门锁信号",
                 门锁9 := "输入"."4号梯9楼层门锁信号",
                 门锁10 := "输入"."4号梯10楼层门锁信号",
                 上下平层同时为1 => "中间变量1".上下平层同时为1梯4,
                 当前楼层数 => "中间变量1"."4号梯当前楼层数",
                 分配当前楼层数 => "中间变量2"."4号梯当前楼层数",
                 正确当前楼层 => "中间变量1"."4号梯正确楼层数");
   END_IF;
END_REGION

REGION Network 6
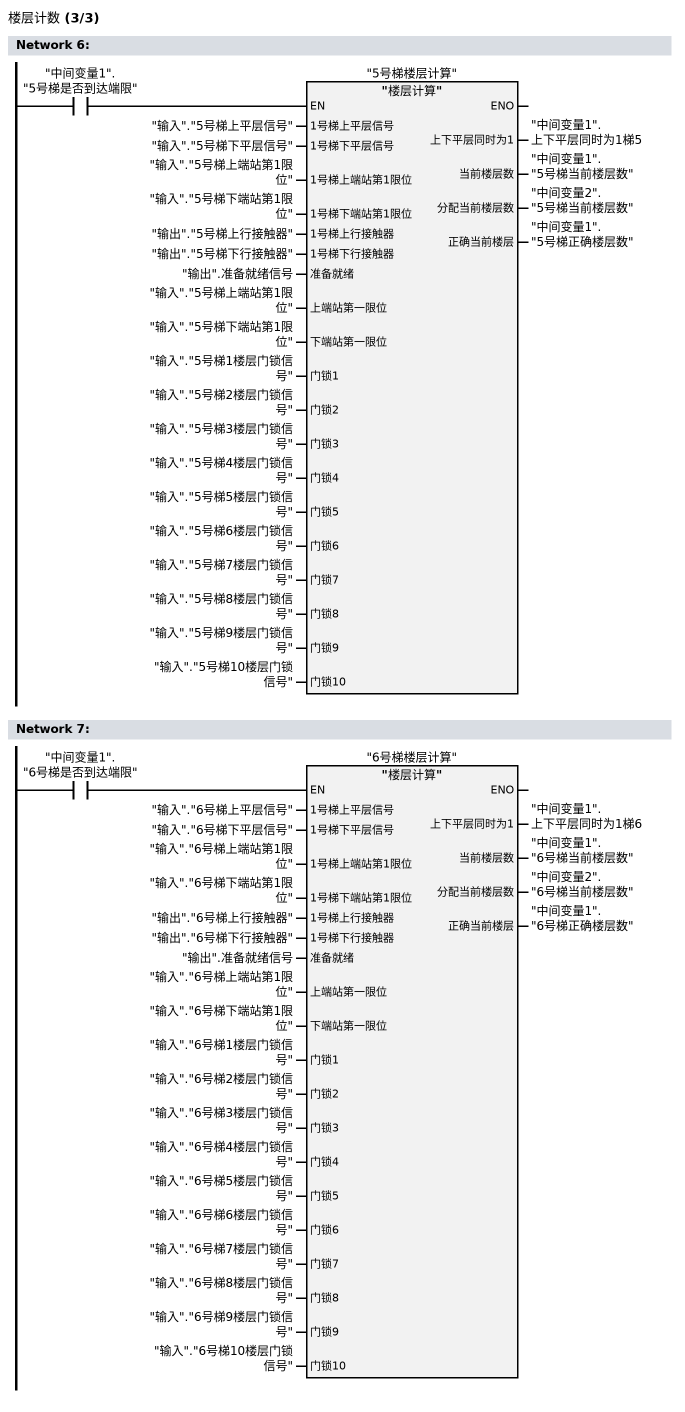
   RUNG wire#powerrail
      Contact( "中间变量1"."5号梯是否到达端限" )
      "5号梯楼层计算"("1号梯上平层信号" := "输入"."5号梯上平层信号", "1号梯下平层信号" := "输入"."5号梯下平层信号", "1号梯上端站第1限位" := "输入"."5号梯上端站第1限位", "1号梯下端站第1限位" := "输入"."5号梯下端站第1限位", "1号梯上行接触器" := "输出"."5号梯上行接触器", "1号梯下行接触器" := "输出"."5号梯下行接触器", 准备就绪 := "输出".准备就绪信号, 上端站第一限位 := "输入"."5号梯上端站第1限位", 下端站第一限位 := "输入"."5号梯下端站第1限位", 门锁1 := "输入"."5号梯1楼层门锁信号", 门锁2 := "输入"."5号梯2楼层门锁信号", 门锁3 := "输入"."5号梯3楼层门锁信号", 门锁4 := "输入"."5号梯4楼层门锁信号", 门锁5 := "输入"."5号梯5楼层门锁信号", 门锁6 := "输入"."5号梯6楼层门锁信号", 门锁7 := "输入"."5号梯7楼层门锁信号", 门锁8 := "输入"."5号梯8楼层门锁信号", 门锁9 := "输入"."5号梯9楼层门锁信号", 门锁10 := "输入"."5号梯10楼层门锁信号", 上下平层同时为1 => "中间变量1".上下平层同时为1梯5, 当前楼层数 => "中间变量1"."5号梯当前楼层数", 分配当前楼层数 => "中间变量2"."5号梯当前楼层数", 正确当前楼层 => "中间变量1"."5号梯正确楼层数")
   END_RUNG
   // the same network as SCL:
   IF "中间变量1"."5号梯是否到达端限" THEN
       "5号梯楼层计算"("1号梯上平层信号" := "输入"."5号梯上平层信号",   // "楼层计算"
                 "1号梯下平层信号" := "输入"."5号梯下平层信号",
                 "1号梯上端站第1限位" := "输入"."5号梯上端站第1限位",
                 "1号梯下端站第1限位" := "输入"."5号梯下端站第1限位",
                 "1号梯上行接触器" := "输出"."5号梯上行接触器",
                 "1号梯下行接触器" := "输出"."5号梯下行接触器",
                 准备就绪 := "输出".准备就绪信号,
                 上端站第一限位 := "输入"."5号梯上端站第1限位",
                 下端站第一限位 := "输入"."5号梯下端站第1限位",
                 门锁1 := "输入"."5号梯1楼层门锁信号",
                 门锁2 := "输入"."5号梯2楼层门锁信号",
                 门锁3 := "输入"."5号梯3楼层门锁信号",
                 门锁4 := "输入"."5号梯4楼层门锁信号",
                 门锁5 := "输入"."5号梯5楼层门锁信号",
                 门锁6 := "输入"."5号梯6楼层门锁信号",
                 门锁7 := "输入"."5号梯7楼层门锁信号",
                 门锁8 := "输入"."5号梯8楼层门锁信号",
                 门锁9 := "输入"."5号梯9楼层门锁信号",
                 门锁10 := "输入"."5号梯10楼层门锁信号",
                 上下平层同时为1 => "中间变量1".上下平层同时为1梯5,
                 当前楼层数 => "中间变量1"."5号梯当前楼层数",
                 分配当前楼层数 => "中间变量2"."5号梯当前楼层数",
                 正确当前楼层 => "中间变量1"."5号梯正确楼层数");
   END_IF;
END_REGION

REGION Network 7
   RUNG wire#powerrail
      Contact( "中间变量1"."6号梯是否到达端限" )
      "6号梯楼层计算"("1号梯上平层信号" := "输入"."6号梯上平层信号", "1号梯下平层信号" := "输入"."6号梯下平层信号", "1号梯上端站第1限位" := "输入"."6号梯上端站第1限位", "1号梯下端站第1限位" := "输入"."6号梯下端站第1限位", "1号梯上行接触器" := "输出"."6号梯上行接触器", "1号梯下行接触器" := "输出"."6号梯下行接触器", 准备就绪 := "输出".准备就绪信号, 上端站第一限位 := "输入"."6号梯上端站第1限位", 下端站第一限位 := "输入"."6号梯下端站第1限位", 门锁1 := "输入"."6号梯1楼层门锁信号", 门锁2 := "输入"."6号梯2楼层门锁信号", 门锁3 := "输入"."6号梯3楼层门锁信号", 门锁4 := "输入"."6号梯4楼层门锁信号", 门锁5 := "输入"."6号梯5楼层门锁信号", 门锁6 := "输入"."6号梯6楼层门锁信号", 门锁7 := "输入"."6号梯7楼层门锁信号", 门锁8 := "输入"."6号梯8楼层门锁信号", 门锁9 := "输入"."6号梯9楼层门锁信号", 门锁10 := "输入"."6号梯10楼层门锁信号", 上下平层同时为1 => "中间变量1".上下平层同时为1梯6, 当前楼层数 => "中间变量1"."6号梯当前楼层数", 分配当前楼层数 => "中间变量2"."6号梯当前楼层数", 正确当前楼层 => "中间变量1"."6号梯正确楼层数")
   END_RUNG
   // the same network as SCL:
   IF "中间变量1"."6号梯是否到达端限" THEN
       "6号梯楼层计算"("1号梯上平层信号" := "输入"."6号梯上平层信号",   // "楼层计算"
                 "1号梯下平层信号" := "输入"."6号梯下平层信号",
                 "1号梯上端站第1限位" := "输入"."6号梯上端站第1限位",
                 "1号梯下端站第1限位" := "输入"."6号梯下端站第1限位",
                 "1号梯上行接触器" := "输出"."6号梯上行接触器",
                 "1号梯下行接触器" := "输出"."6号梯下行接触器",
                 准备就绪 := "输出".准备就绪信号,
                 上端站第一限位 := "输入"."6号梯上端站第1限位",
                 下端站第一限位 := "输入"."6号梯下端站第1限位",
                 门锁1 := "输入"."6号梯1楼层门锁信号",
                 门锁2 := "输入"."6号梯2楼层门锁信号",
                 门锁3 := "输入"."6号梯3楼层门锁信号",
                 门锁4 := "输入"."6号梯4楼层门锁信号",
                 门锁5 := "输入"."6号梯5楼层门锁信号",
                 门锁6 := "输入"."6号梯6楼层门锁信号",
                 门锁7 := "输入"."6号梯7楼层门锁信号",
                 门锁8 := "输入"."6号梯8楼层门锁信号",
                 门锁9 := "输入"."6号梯9楼层门锁信号",
                 门锁10 := "输入"."6号梯10楼层门锁信号",
                 上下平层同时为1 => "中间变量1".上下平层同时为1梯6,
                 当前楼层数 => "中间变量1"."6号梯当前楼层数",
                 分配当前楼层数 => "中间变量2"."6号梯当前楼层数",
                 正确当前楼层 => "中间变量1"."6号梯正确楼层数");
   END_IF;
END_REGION
END_FUNCTION

FUNCTION "优先级" : Void   // FC10, LAD
{ S7_Optimized_Access := 'TRUE' }
VERSION : 0.1
BEGIN

REGION Network 2: 1
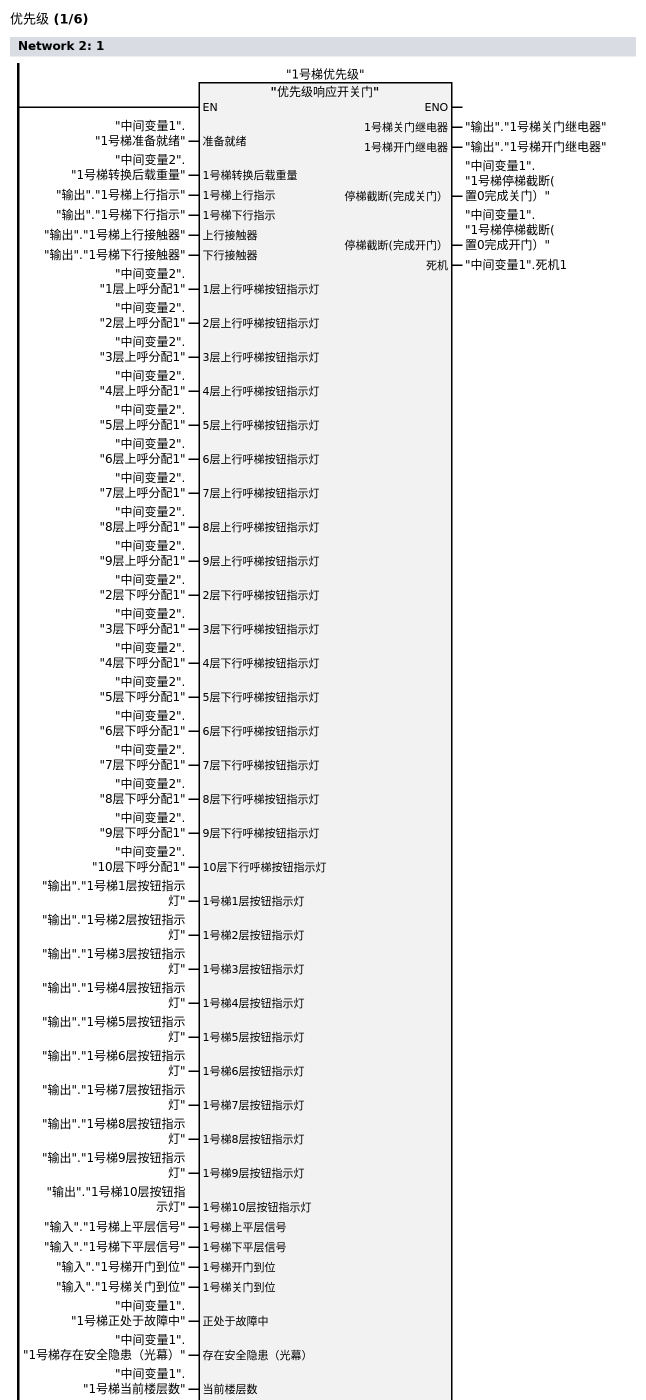
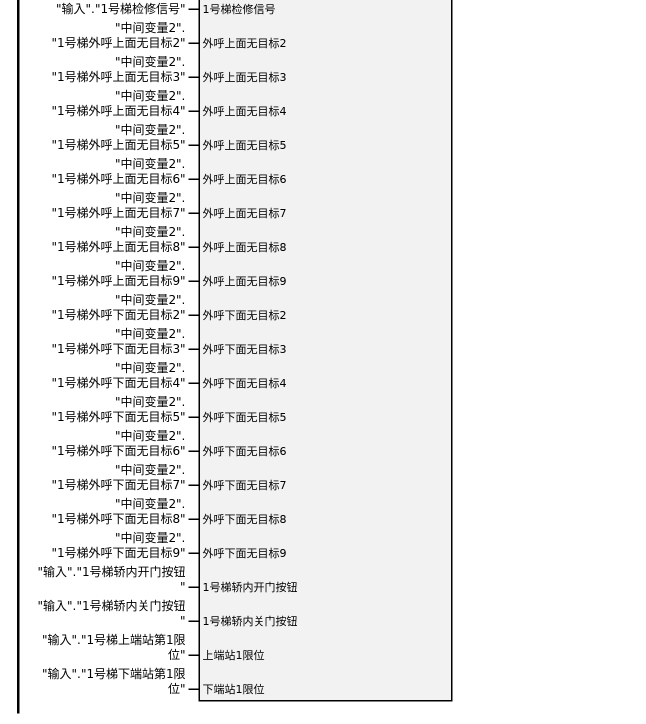
   RUNG wire#powerrail
      "1号梯优先级"(准备就绪 := "中间变量1"."1号梯准备就绪", "1号梯转换后载重量" := "中间变量2"."1号梯转换后载重量", "1号梯上行指示" := "输出"."1号梯上行指示", "1号梯下行指示" := "输出"."1号梯下行指示", 上行接触器 := "输出"."1号梯上行接触器", 下行接触器 := "输出"."1号梯下行接触器", "1层上行呼梯按钮指示灯" := "中间变量2"."1层上呼分配1", "2层上行呼梯按钮指示灯" := "中间变量2"."2层上呼分配1", "3层上行呼梯按钮指示灯" := "中间变量2"."3层上呼分配1", "4层上行呼梯按钮指示灯" := "中间变量2"."4层上呼分配1", "5层上行呼梯按钮指示灯" := "中间变量2"."5层上呼分配1", "6层上行呼梯按钮指示灯" := "中间变量2"."6层上呼分配1", "7层上行呼梯按钮指示灯" := "中间变量2"."7层上呼分配1", "8层上行呼梯按钮指示灯" := "中间变量2"."8层上呼分配1", "9层上行呼梯按钮指示灯" := "中间变量2"."9层上呼分配1", "2层下行呼梯按钮指示灯" := "中间变量2"."2层下呼分配1", "3层下行呼梯按钮指示灯" := "中间变量2"."3层下呼分配1", "4层下行呼梯按钮指示灯" := "中间变量2"."4层下呼分配1", "5层下行呼梯按钮指示灯" := "中间变量2"."5层下呼分配1", "6层下行呼梯按钮指示灯" := "中间变量2"."6层下呼分配1", "7层下行呼梯按钮指示灯" := "中间变量2"."7层下呼分配1", "8层下行呼梯按钮指示灯" := "中间变量2"."8层下呼分配1", "9层下行呼梯按钮指示灯" := "中间变量2"."9层下呼分配1", "10层下行呼梯按钮指示灯" := "中间变量2"."10层下呼分配1", "1号梯1层按钮指示灯" := "输出"."1号梯1层按钮指示灯", "1号梯2层按钮指示灯" := "输出"."1号梯2层按钮指示灯", "1号梯3层按钮指示灯" := "输出"."1号梯3层按钮指示灯", "1号梯4层按钮指示灯" := "输出"."1号梯4层按钮指示灯", "1号梯5层按钮指示灯" := "输出"."1号梯5层按钮指示灯", "1号梯6层按钮指示灯" := "输出"."1号梯6层按钮指示灯", "1号梯7层按钮指示灯" := "输出"."1号梯7层按钮指示灯", "1号梯8层按钮指示灯" := "输出"."1号梯8层按钮指示灯", "1号梯9层按钮指示灯" := "输出"."1号梯9层按钮指示灯", "1号梯10层按钮指示灯" := "输出"."1号梯10层按钮指示灯", "1号梯上平层信号" := "输入"."1号梯上平层信号", "1号梯下平层信号" := "输入"."1号梯下平层信号", "1号梯开门到位" := "输入"."1号梯开门到位", "1号梯关门到位" := "输入"."1号梯关门到位", 正处于故障中 := "中间变量1"."1号梯正处于故障中", "存在安全隐患（光幕）" := "中间变量1"."1号梯存在安全隐患（光幕）", 当前楼层数 := "中间变量1"."1号梯当前楼层数", "1号梯检修信号" := "输入"."1号梯检修信号", 外呼上面无目标2 := "中间变量2"."1号梯外呼上面无目标2", 外呼上面无目标3 := "中间变量2"."1号梯外呼上面无目标3", 外呼上面无目标4 := "中间变量2"."1号梯外呼上面无目标4", 外呼上面无目标5 := "中间变量2"."1号梯外呼上面无目标5", 外呼上面无目标6 := "中间变量2"."1号梯外呼上面无目标6", 外呼上面无目标7 := "中间变量2"."1号梯外呼上面无目标7", 外呼上面无目标8 := "中间变量2"."1号梯外呼上面无目标8", 外呼上面无目标9 := "中间变量2"."1号梯外呼上面无目标9", 外呼下面无目标2 := "中间变量2"."1号梯外呼下面无目标2", 外呼下面无目标3 := "中间变量2"."1号梯外呼下面无目标3", 外呼下面无目标4 := "中间变量2"."1号梯外呼下面无目标4", 外呼下面无目标5 := "中间变量2"."1号梯外呼下面无目标5", 外呼下面无目标6 := "中间变量2"."1号梯外呼下面无目标6", 外呼下面无目标7 := "中间变量2"."1号梯外呼下面无目标7", 外呼下面无目标8 := "中间变量2"."1号梯外呼下面无目标8", 外呼下面无目标9 := "中间变量2"."1号梯外呼下面无目标9", "1号梯轿内开门按钮" := "输入"."1号梯轿内开门按钮", "1号梯轿内关门按钮" := "输入"."1号梯轿内关门按钮", 上端站1限位 := "输入"."1号梯上端站第1限位", 下端站1限位 := "输入"."1号梯下端站第1限位", "1号梯关门继电器" => "输出"."1号梯关门继电器", "1号梯开门继电器" => "输出"."1号梯开门继电器", "停梯截断(完成关门）" => "中间变量1"."1号梯停梯截断(置0完成关门）", "停梯截断(完成开门）" => "中间变量1"."1号梯停梯截断(置0完成开门）", 死机 => "中间变量1".死机1)
   END_RUNG
   // the same network as SCL:
   "1号梯优先级"(准备就绪 := "中间变量1"."1号梯准备就绪",   // "优先级响应开关门"
            "1号梯转换后载重量" := "中间变量2"."1号梯转换后载重量",
            "1号梯上行指示" := "输出"."1号梯上行指示",
            "1号梯下行指示" := "输出"."1号梯下行指示",
            上行接触器 := "输出"."1号梯上行接触器",
            下行接触器 := "输出"."1号梯下行接触器",
            "1层上行呼梯按钮指示灯" := "中间变量2"."1层上呼分配1",
            "2层上行呼梯按钮指示灯" := "中间变量2"."2层上呼分配1",
            "3层上行呼梯按钮指示灯" := "中间变量2"."3层上呼分配1",
            "4层上行呼梯按钮指示灯" := "中间变量2"."4层上呼分配1",
            "5层上行呼梯按钮指示灯" := "中间变量2"."5层上呼分配1",
            "6层上行呼梯按钮指示灯" := "中间变量2"."6层上呼分配1",
            "7层上行呼梯按钮指示灯" := "中间变量2"."7层上呼分配1",
            "8层上行呼梯按钮指示灯" := "中间变量2"."8层上呼分配1",
            "9层上行呼梯按钮指示灯" := "中间变量2"."9层上呼分配1",
            "2层下行呼梯按钮指示灯" := "中间变量2"."2层下呼分配1",
            "3层下行呼梯按钮指示灯" := "中间变量2"."3层下呼分配1",
            "4层下行呼梯按钮指示灯" := "中间变量2"."4层下呼分配1",
            "5层下行呼梯按钮指示灯" := "中间变量2"."5层下呼分配1",
            "6层下行呼梯按钮指示灯" := "中间变量2"."6层下呼分配1",
            "7层下行呼梯按钮指示灯" := "中间变量2"."7层下呼分配1",
            "8层下行呼梯按钮指示灯" := "中间变量2"."8层下呼分配1",
            "9层下行呼梯按钮指示灯" := "中间变量2"."9层下呼分配1",
            "10层下行呼梯按钮指示灯" := "中间变量2"."10层下呼分配1",
            "1号梯1层按钮指示灯" := "输出"."1号梯1层按钮指示灯",
            "1号梯2层按钮指示灯" := "输出"."1号梯2层按钮指示灯",
            "1号梯3层按钮指示灯" := "输出"."1号梯3层按钮指示灯",
            "1号梯4层按钮指示灯" := "输出"."1号梯4层按钮指示灯",
            "1号梯5层按钮指示灯" := "输出"."1号梯5层按钮指示灯",
            "1号梯6层按钮指示灯" := "输出"."1号梯6层按钮指示灯",
            "1号梯7层按钮指示灯" := "输出"."1号梯7层按钮指示灯",
            "1号梯8层按钮指示灯" := "输出"."1号梯8层按钮指示灯",
            "1号梯9层按钮指示灯" := "输出"."1号梯9层按钮指示灯",
            "1号梯10层按钮指示灯" := "输出"."1号梯10层按钮指示灯",
            "1号梯上平层信号" := "输入"."1号梯上平层信号",
            "1号梯下平层信号" := "输入"."1号梯下平层信号",
            "1号梯开门到位" := "输入"."1号梯开门到位",
            "1号梯关门到位" := "输入"."1号梯关门到位",
            正处于故障中 := "中间变量1"."1号梯正处于故障中",
            "存在安全隐患（光幕）" := "中间变量1"."1号梯存在安全隐患（光幕）",
            当前楼层数 := "中间变量1"."1号梯当前楼层数",
            "1号梯检修信号" := "输入"."1号梯检修信号",
            外呼上面无目标2 := "中间变量2"."1号梯外呼上面无目标2",
            外呼上面无目标3 := "中间变量2"."1号梯外呼上面无目标3",
            外呼上面无目标4 := "中间变量2"."1号梯外呼上面无目标4",
            外呼上面无目标5 := "中间变量2"."1号梯外呼上面无目标5",
            外呼上面无目标6 := "中间变量2"."1号梯外呼上面无目标6",
            外呼上面无目标7 := "中间变量2"."1号梯外呼上面无目标7",
            外呼上面无目标8 := "中间变量2"."1号梯外呼上面无目标8",
            外呼上面无目标9 := "中间变量2"."1号梯外呼上面无目标9",
            外呼下面无目标2 := "中间变量2"."1号梯外呼下面无目标2",
            外呼下面无目标3 := "中间变量2"."1号梯外呼下面无目标3",
            外呼下面无目标4 := "中间变量2"."1号梯外呼下面无目标4",
            外呼下面无目标5 := "中间变量2"."1号梯外呼下面无目标5",
            外呼下面无目标6 := "中间变量2"."1号梯外呼下面无目标6",
            外呼下面无目标7 := "中间变量2"."1号梯外呼下面无目标7",
            外呼下面无目标8 := "中间变量2"."1号梯外呼下面无目标8",
            外呼下面无目标9 := "中间变量2"."1号梯外呼下面无目标9",
            "1号梯轿内开门按钮" := "输入"."1号梯轿内开门按钮",
            "1号梯轿内关门按钮" := "输入"."1号梯轿内关门按钮",
            上端站1限位 := "输入"."1号梯上端站第1限位",
            下端站1限位 := "输入"."1号梯下端站第1限位",
            "1号梯关门继电器" => "输出"."1号梯关门继电器",
            "1号梯开门继电器" => "输出"."1号梯开门继电器",
            "停梯截断(完成关门）" => "中间变量1"."1号梯停梯截断(置0完成关门）",
            "停梯截断(完成开门）" => "中间变量1"."1号梯停梯截断(置0完成开门）",
            死机 => "中间变量1".死机1);
END_REGION

REGION Network 3: 2
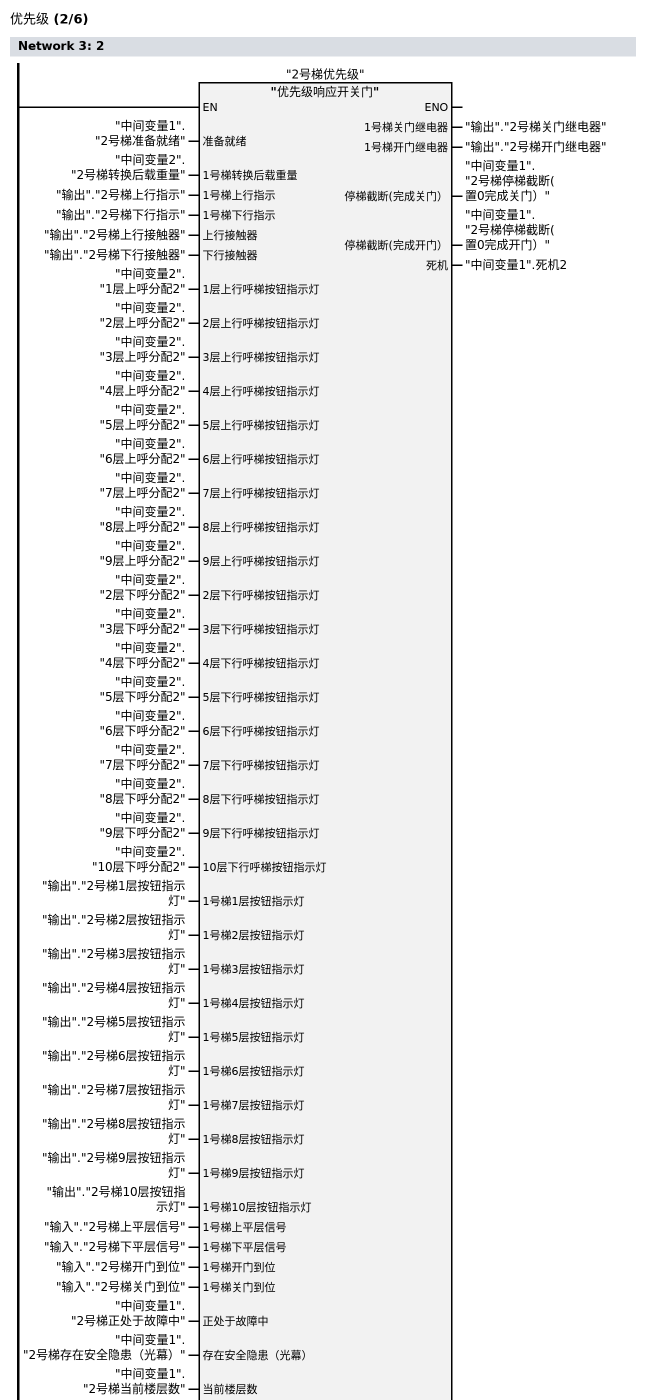
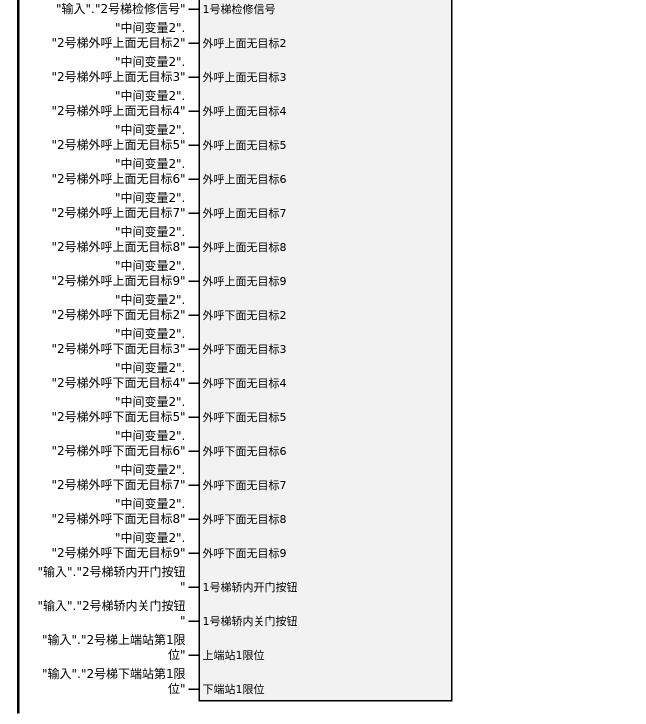
   RUNG wire#powerrail
      "2号梯优先级"(准备就绪 := "中间变量1"."2号梯准备就绪", "1号梯转换后载重量" := "中间变量2"."2号梯转换后载重量", "1号梯上行指示" := "输出"."2号梯上行指示", "1号梯下行指示" := "输出"."2号梯下行指示", 上行接触器 := "输出"."2号梯上行接触器", 下行接触器 := "输出"."2号梯下行接触器", "1层上行呼梯按钮指示灯" := "中间变量2"."1层上呼分配2", "2层上行呼梯按钮指示灯" := "中间变量2"."2层上呼分配2", "3层上行呼梯按钮指示灯" := "中间变量2"."3层上呼分配2", "4层上行呼梯按钮指示灯" := "中间变量2"."4层上呼分配2", "5层上行呼梯按钮指示灯" := "中间变量2"."5层上呼分配2", "6层上行呼梯按钮指示灯" := "中间变量2"."6层上呼分配2", "7层上行呼梯按钮指示灯" := "中间变量2"."7层上呼分配2", "8层上行呼梯按钮指示灯" := "中间变量2"."8层上呼分配2", "9层上行呼梯按钮指示灯" := "中间变量2"."9层上呼分配2", "2层下行呼梯按钮指示灯" := "中间变量2"."2层下呼分配2", "3层下行呼梯按钮指示灯" := "中间变量2"."3层下呼分配2", "4层下行呼梯按钮指示灯" := "中间变量2"."4层下呼分配2", "5层下行呼梯按钮指示灯" := "中间变量2"."5层下呼分配2", "6层下行呼梯按钮指示灯" := "中间变量2"."6层下呼分配2", "7层下行呼梯按钮指示灯" := "中间变量2"."7层下呼分配2", "8层下行呼梯按钮指示灯" := "中间变量2"."8层下呼分配2", "9层下行呼梯按钮指示灯" := "中间变量2"."9层下呼分配2", "10层下行呼梯按钮指示灯" := "中间变量2"."10层下呼分配2", "1号梯1层按钮指示灯" := "输出"."2号梯1层按钮指示灯", "1号梯2层按钮指示灯" := "输出"."2号梯2层按钮指示灯", "1号梯3层按钮指示灯" := "输出"."2号梯3层按钮指示灯", "1号梯4层按钮指示灯" := "输出"."2号梯4层按钮指示灯", "1号梯5层按钮指示灯" := "输出"."2号梯5层按钮指示灯", "1号梯6层按钮指示灯" := "输出"."2号梯6层按钮指示灯", "1号梯7层按钮指示灯" := "输出"."2号梯7层按钮指示灯", "1号梯8层按钮指示灯" := "输出"."2号梯8层按钮指示灯", "1号梯9层按钮指示灯" := "输出"."2号梯9层按钮指示灯", "1号梯10层按钮指示灯" := "输出"."2号梯10层按钮指示灯", "1号梯上平层信号" := "输入"."2号梯上平层信号", "1号梯下平层信号" := "输入"."2号梯下平层信号", "1号梯开门到位" := "输入"."2号梯开门到位", "1号梯关门到位" := "输入"."2号梯关门到位", 正处于故障中 := "中间变量1"."2号梯正处于故障中", "存在安全隐患（光幕）" := "中间变量1"."2号梯存在安全隐患（光幕）", 当前楼层数 := "中间变量1"."2号梯当前楼层数", "1号梯检修信号" := "输入"."2号梯检修信号", 外呼上面无目标2 := "中间变量2"."2号梯外呼上面无目标2", 外呼上面无目标3 := "中间变量2"."2号梯外呼上面无目标3", 外呼上面无目标4 := "中间变量2"."2号梯外呼上面无目标4", 外呼上面无目标5 := "中间变量2"."2号梯外呼上面无目标5", 外呼上面无目标6 := "中间变量2"."2号梯外呼上面无目标6", 外呼上面无目标7 := "中间变量2"."2号梯外呼上面无目标7", 外呼上面无目标8 := "中间变量2"."2号梯外呼上面无目标8", 外呼上面无目标9 := "中间变量2"."2号梯外呼上面无目标9", 外呼下面无目标2 := "中间变量2"."2号梯外呼下面无目标2", 外呼下面无目标3 := "中间变量2"."2号梯外呼下面无目标3", 外呼下面无目标4 := "中间变量2"."2号梯外呼下面无目标4", 外呼下面无目标5 := "中间变量2"."2号梯外呼下面无目标5", 外呼下面无目标6 := "中间变量2"."2号梯外呼下面无目标6", 外呼下面无目标7 := "中间变量2"."2号梯外呼下面无目标7", 外呼下面无目标8 := "中间变量2"."2号梯外呼下面无目标8", 外呼下面无目标9 := "中间变量2"."2号梯外呼下面无目标9", "1号梯轿内开门按钮" := "输入"."2号梯轿内开门按钮", "1号梯轿内关门按钮" := "输入"."2号梯轿内关门按钮", 上端站1限位 := "输入"."2号梯上端站第1限位", 下端站1限位 := "输入"."2号梯下端站第1限位", "1号梯关门继电器" => "输出"."2号梯关门继电器", "1号梯开门继电器" => "输出"."2号梯开门继电器", "停梯截断(完成关门）" => "中间变量1"."2号梯停梯截断(置0完成关门）", "停梯截断(完成开门）" => "中间变量1"."2号梯停梯截断(置0完成开门）", 死机 => "中间变量1".死机2)
   END_RUNG
   // the same network as SCL:
   "2号梯优先级"(准备就绪 := "中间变量1"."2号梯准备就绪",   // "优先级响应开关门"
            "1号梯转换后载重量" := "中间变量2"."2号梯转换后载重量",
            "1号梯上行指示" := "输出"."2号梯上行指示",
            "1号梯下行指示" := "输出"."2号梯下行指示",
            上行接触器 := "输出"."2号梯上行接触器",
            下行接触器 := "输出"."2号梯下行接触器",
            "1层上行呼梯按钮指示灯" := "中间变量2"."1层上呼分配2",
            "2层上行呼梯按钮指示灯" := "中间变量2"."2层上呼分配2",
            "3层上行呼梯按钮指示灯" := "中间变量2"."3层上呼分配2",
            "4层上行呼梯按钮指示灯" := "中间变量2"."4层上呼分配2",
            "5层上行呼梯按钮指示灯" := "中间变量2"."5层上呼分配2",
            "6层上行呼梯按钮指示灯" := "中间变量2"."6层上呼分配2",
            "7层上行呼梯按钮指示灯" := "中间变量2"."7层上呼分配2",
            "8层上行呼梯按钮指示灯" := "中间变量2"."8层上呼分配2",
            "9层上行呼梯按钮指示灯" := "中间变量2"."9层上呼分配2",
            "2层下行呼梯按钮指示灯" := "中间变量2"."2层下呼分配2",
            "3层下行呼梯按钮指示灯" := "中间变量2"."3层下呼分配2",
            "4层下行呼梯按钮指示灯" := "中间变量2"."4层下呼分配2",
            "5层下行呼梯按钮指示灯" := "中间变量2"."5层下呼分配2",
            "6层下行呼梯按钮指示灯" := "中间变量2"."6层下呼分配2",
            "7层下行呼梯按钮指示灯" := "中间变量2"."7层下呼分配2",
            "8层下行呼梯按钮指示灯" := "中间变量2"."8层下呼分配2",
            "9层下行呼梯按钮指示灯" := "中间变量2"."9层下呼分配2",
            "10层下行呼梯按钮指示灯" := "中间变量2"."10层下呼分配2",
            "1号梯1层按钮指示灯" := "输出"."2号梯1层按钮指示灯",
            "1号梯2层按钮指示灯" := "输出"."2号梯2层按钮指示灯",
            "1号梯3层按钮指示灯" := "输出"."2号梯3层按钮指示灯",
            "1号梯4层按钮指示灯" := "输出"."2号梯4层按钮指示灯",
            "1号梯5层按钮指示灯" := "输出"."2号梯5层按钮指示灯",
            "1号梯6层按钮指示灯" := "输出"."2号梯6层按钮指示灯",
            "1号梯7层按钮指示灯" := "输出"."2号梯7层按钮指示灯",
            "1号梯8层按钮指示灯" := "输出"."2号梯8层按钮指示灯",
            "1号梯9层按钮指示灯" := "输出"."2号梯9层按钮指示灯",
            "1号梯10层按钮指示灯" := "输出"."2号梯10层按钮指示灯",
            "1号梯上平层信号" := "输入"."2号梯上平层信号",
            "1号梯下平层信号" := "输入"."2号梯下平层信号",
            "1号梯开门到位" := "输入"."2号梯开门到位",
            "1号梯关门到位" := "输入"."2号梯关门到位",
            正处于故障中 := "中间变量1"."2号梯正处于故障中",
            "存在安全隐患（光幕）" := "中间变量1"."2号梯存在安全隐患（光幕）",
            当前楼层数 := "中间变量1"."2号梯当前楼层数",
            "1号梯检修信号" := "输入"."2号梯检修信号",
            外呼上面无目标2 := "中间变量2"."2号梯外呼上面无目标2",
            外呼上面无目标3 := "中间变量2"."2号梯外呼上面无目标3",
            外呼上面无目标4 := "中间变量2"."2号梯外呼上面无目标4",
            外呼上面无目标5 := "中间变量2"."2号梯外呼上面无目标5",
            外呼上面无目标6 := "中间变量2"."2号梯外呼上面无目标6",
            外呼上面无目标7 := "中间变量2"."2号梯外呼上面无目标7",
            外呼上面无目标8 := "中间变量2"."2号梯外呼上面无目标8",
            外呼上面无目标9 := "中间变量2"."2号梯外呼上面无目标9",
            外呼下面无目标2 := "中间变量2"."2号梯外呼下面无目标2",
            外呼下面无目标3 := "中间变量2"."2号梯外呼下面无目标3",
            外呼下面无目标4 := "中间变量2"."2号梯外呼下面无目标4",
            外呼下面无目标5 := "中间变量2"."2号梯外呼下面无目标5",
            外呼下面无目标6 := "中间变量2"."2号梯外呼下面无目标6",
            外呼下面无目标7 := "中间变量2"."2号梯外呼下面无目标7",
            外呼下面无目标8 := "中间变量2"."2号梯外呼下面无目标8",
            外呼下面无目标9 := "中间变量2"."2号梯外呼下面无目标9",
            "1号梯轿内开门按钮" := "输入"."2号梯轿内开门按钮",
            "1号梯轿内关门按钮" := "输入"."2号梯轿内关门按钮",
            上端站1限位 := "输入"."2号梯上端站第1限位",
            下端站1限位 := "输入"."2号梯下端站第1限位",
            "1号梯关门继电器" => "输出"."2号梯关门继电器",
            "1号梯开门继电器" => "输出"."2号梯开门继电器",
            "停梯截断(完成关门）" => "中间变量1"."2号梯停梯截断(置0完成关门）",
            "停梯截断(完成开门）" => "中间变量1"."2号梯停梯截断(置0完成开门）",
            死机 => "中间变量1".死机2);
END_REGION

REGION Network 4: 3
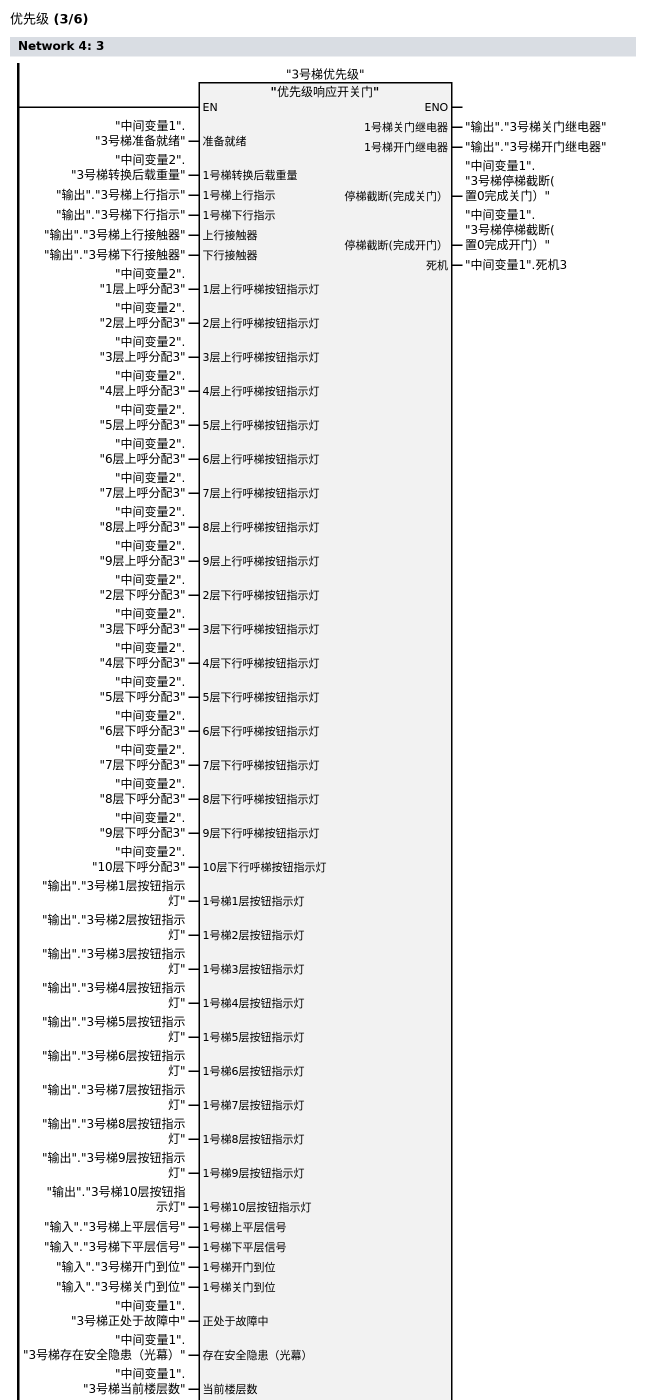
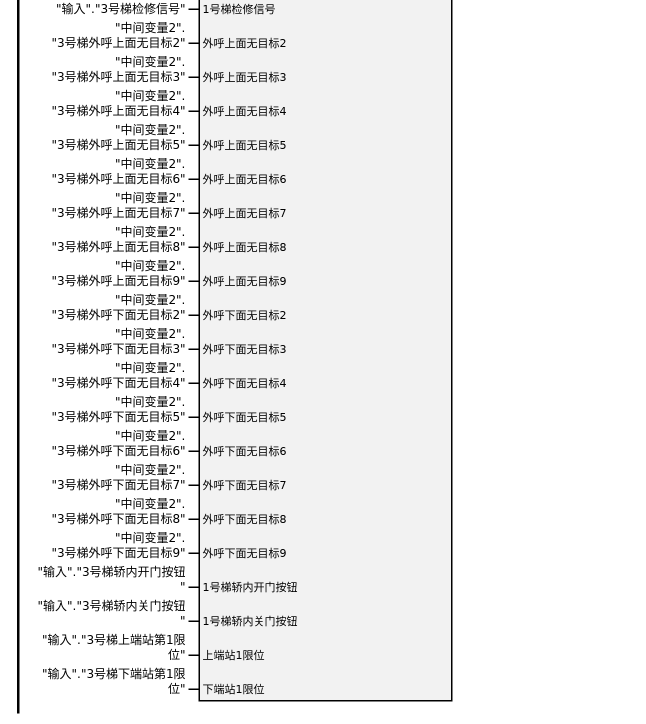
   RUNG wire#powerrail
      "3号梯优先级"(准备就绪 := "中间变量1"."3号梯准备就绪", "1号梯转换后载重量" := "中间变量2"."3号梯转换后载重量", "1号梯上行指示" := "输出"."3号梯上行指示", "1号梯下行指示" := "输出"."3号梯下行指示", 上行接触器 := "输出"."3号梯上行接触器", 下行接触器 := "输出"."3号梯下行接触器", "1层上行呼梯按钮指示灯" := "中间变量2"."1层上呼分配3", "2层上行呼梯按钮指示灯" := "中间变量2"."2层上呼分配3", "3层上行呼梯按钮指示灯" := "中间变量2"."3层上呼分配3", "4层上行呼梯按钮指示灯" := "中间变量2"."4层上呼分配3", "5层上行呼梯按钮指示灯" := "中间变量2"."5层上呼分配3", "6层上行呼梯按钮指示灯" := "中间变量2"."6层上呼分配3", "7层上行呼梯按钮指示灯" := "中间变量2"."7层上呼分配3", "8层上行呼梯按钮指示灯" := "中间变量2"."8层上呼分配3", "9层上行呼梯按钮指示灯" := "中间变量2"."9层上呼分配3", "2层下行呼梯按钮指示灯" := "中间变量2"."2层下呼分配3", "3层下行呼梯按钮指示灯" := "中间变量2"."3层下呼分配3", "4层下行呼梯按钮指示灯" := "中间变量2"."4层下呼分配3", "5层下行呼梯按钮指示灯" := "中间变量2"."5层下呼分配3", "6层下行呼梯按钮指示灯" := "中间变量2"."6层下呼分配3", "7层下行呼梯按钮指示灯" := "中间变量2"."7层下呼分配3", "8层下行呼梯按钮指示灯" := "中间变量2"."8层下呼分配3", "9层下行呼梯按钮指示灯" := "中间变量2"."9层下呼分配3", "10层下行呼梯按钮指示灯" := "中间变量2"."10层下呼分配3", "1号梯1层按钮指示灯" := "输出"."3号梯1层按钮指示灯", "1号梯2层按钮指示灯" := "输出"."3号梯2层按钮指示灯", "1号梯3层按钮指示灯" := "输出"."3号梯3层按钮指示灯", "1号梯4层按钮指示灯" := "输出"."3号梯4层按钮指示灯", "1号梯5层按钮指示灯" := "输出"."3号梯5层按钮指示灯", "1号梯6层按钮指示灯" := "输出"."3号梯6层按钮指示灯", "1号梯7层按钮指示灯" := "输出"."3号梯7层按钮指示灯", "1号梯8层按钮指示灯" := "输出"."3号梯8层按钮指示灯", "1号梯9层按钮指示灯" := "输出"."3号梯9层按钮指示灯", "1号梯10层按钮指示灯" := "输出"."3号梯10层按钮指示灯", "1号梯上平层信号" := "输入"."3号梯上平层信号", "1号梯下平层信号" := "输入"."3号梯下平层信号", "1号梯开门到位" := "输入"."3号梯开门到位", "1号梯关门到位" := "输入"."3号梯关门到位", 正处于故障中 := "中间变量1"."3号梯正处于故障中", "存在安全隐患（光幕）" := "中间变量1"."3号梯存在安全隐患（光幕）", 当前楼层数 := "中间变量1"."3号梯当前楼层数", "1号梯检修信号" := "输入"."3号梯检修信号", 外呼上面无目标2 := "中间变量2"."3号梯外呼上面无目标2", 外呼上面无目标3 := "中间变量2"."3号梯外呼上面无目标3", 外呼上面无目标4 := "中间变量2"."3号梯外呼上面无目标4", 外呼上面无目标5 := "中间变量2"."3号梯外呼上面无目标5", 外呼上面无目标6 := "中间变量2"."3号梯外呼上面无目标6", 外呼上面无目标7 := "中间变量2"."3号梯外呼上面无目标7", 外呼上面无目标8 := "中间变量2"."3号梯外呼上面无目标8", 外呼上面无目标9 := "中间变量2"."3号梯外呼上面无目标9", 外呼下面无目标2 := "中间变量2"."3号梯外呼下面无目标2", 外呼下面无目标3 := "中间变量2"."3号梯外呼下面无目标3", 外呼下面无目标4 := "中间变量2"."3号梯外呼下面无目标4", 外呼下面无目标5 := "中间变量2"."3号梯外呼下面无目标5", 外呼下面无目标6 := "中间变量2"."3号梯外呼下面无目标6", 外呼下面无目标7 := "中间变量2"."3号梯外呼下面无目标7", 外呼下面无目标8 := "中间变量2"."3号梯外呼下面无目标8", 外呼下面无目标9 := "中间变量2"."3号梯外呼下面无目标9", "1号梯轿内开门按钮" := "输入"."3号梯轿内开门按钮", "1号梯轿内关门按钮" := "输入"."3号梯轿内关门按钮", 上端站1限位 := "输入"."3号梯上端站第1限位", 下端站1限位 := "输入"."3号梯下端站第1限位", "1号梯关门继电器" => "输出"."3号梯关门继电器", "1号梯开门继电器" => "输出"."3号梯开门继电器", "停梯截断(完成关门）" => "中间变量1"."3号梯停梯截断(置0完成关门）", "停梯截断(完成开门）" => "中间变量1"."3号梯停梯截断(置0完成开门）", 死机 => "中间变量1".死机3)
   END_RUNG
   // the same network as SCL:
   "3号梯优先级"(准备就绪 := "中间变量1"."3号梯准备就绪",   // "优先级响应开关门"
            "1号梯转换后载重量" := "中间变量2"."3号梯转换后载重量",
            "1号梯上行指示" := "输出"."3号梯上行指示",
            "1号梯下行指示" := "输出"."3号梯下行指示",
            上行接触器 := "输出"."3号梯上行接触器",
            下行接触器 := "输出"."3号梯下行接触器",
            "1层上行呼梯按钮指示灯" := "中间变量2"."1层上呼分配3",
            "2层上行呼梯按钮指示灯" := "中间变量2"."2层上呼分配3",
            "3层上行呼梯按钮指示灯" := "中间变量2"."3层上呼分配3",
            "4层上行呼梯按钮指示灯" := "中间变量2"."4层上呼分配3",
            "5层上行呼梯按钮指示灯" := "中间变量2"."5层上呼分配3",
            "6层上行呼梯按钮指示灯" := "中间变量2"."6层上呼分配3",
            "7层上行呼梯按钮指示灯" := "中间变量2"."7层上呼分配3",
            "8层上行呼梯按钮指示灯" := "中间变量2"."8层上呼分配3",
            "9层上行呼梯按钮指示灯" := "中间变量2"."9层上呼分配3",
            "2层下行呼梯按钮指示灯" := "中间变量2"."2层下呼分配3",
            "3层下行呼梯按钮指示灯" := "中间变量2"."3层下呼分配3",
            "4层下行呼梯按钮指示灯" := "中间变量2"."4层下呼分配3",
            "5层下行呼梯按钮指示灯" := "中间变量2"."5层下呼分配3",
            "6层下行呼梯按钮指示灯" := "中间变量2"."6层下呼分配3",
            "7层下行呼梯按钮指示灯" := "中间变量2"."7层下呼分配3",
            "8层下行呼梯按钮指示灯" := "中间变量2"."8层下呼分配3",
            "9层下行呼梯按钮指示灯" := "中间变量2"."9层下呼分配3",
            "10层下行呼梯按钮指示灯" := "中间变量2"."10层下呼分配3",
            "1号梯1层按钮指示灯" := "输出"."3号梯1层按钮指示灯",
            "1号梯2层按钮指示灯" := "输出"."3号梯2层按钮指示灯",
            "1号梯3层按钮指示灯" := "输出"."3号梯3层按钮指示灯",
            "1号梯4层按钮指示灯" := "输出"."3号梯4层按钮指示灯",
            "1号梯5层按钮指示灯" := "输出"."3号梯5层按钮指示灯",
            "1号梯6层按钮指示灯" := "输出"."3号梯6层按钮指示灯",
            "1号梯7层按钮指示灯" := "输出"."3号梯7层按钮指示灯",
            "1号梯8层按钮指示灯" := "输出"."3号梯8层按钮指示灯",
            "1号梯9层按钮指示灯" := "输出"."3号梯9层按钮指示灯",
            "1号梯10层按钮指示灯" := "输出"."3号梯10层按钮指示灯",
            "1号梯上平层信号" := "输入"."3号梯上平层信号",
            "1号梯下平层信号" := "输入"."3号梯下平层信号",
            "1号梯开门到位" := "输入"."3号梯开门到位",
            "1号梯关门到位" := "输入"."3号梯关门到位",
            正处于故障中 := "中间变量1"."3号梯正处于故障中",
            "存在安全隐患（光幕）" := "中间变量1"."3号梯存在安全隐患（光幕）",
            当前楼层数 := "中间变量1"."3号梯当前楼层数",
            "1号梯检修信号" := "输入"."3号梯检修信号",
            外呼上面无目标2 := "中间变量2"."3号梯外呼上面无目标2",
            外呼上面无目标3 := "中间变量2"."3号梯外呼上面无目标3",
            外呼上面无目标4 := "中间变量2"."3号梯外呼上面无目标4",
            外呼上面无目标5 := "中间变量2"."3号梯外呼上面无目标5",
            外呼上面无目标6 := "中间变量2"."3号梯外呼上面无目标6",
            外呼上面无目标7 := "中间变量2"."3号梯外呼上面无目标7",
            外呼上面无目标8 := "中间变量2"."3号梯外呼上面无目标8",
            外呼上面无目标9 := "中间变量2"."3号梯外呼上面无目标9",
            外呼下面无目标2 := "中间变量2"."3号梯外呼下面无目标2",
            外呼下面无目标3 := "中间变量2"."3号梯外呼下面无目标3",
            外呼下面无目标4 := "中间变量2"."3号梯外呼下面无目标4",
            外呼下面无目标5 := "中间变量2"."3号梯外呼下面无目标5",
            外呼下面无目标6 := "中间变量2"."3号梯外呼下面无目标6",
            外呼下面无目标7 := "中间变量2"."3号梯外呼下面无目标7",
            外呼下面无目标8 := "中间变量2"."3号梯外呼下面无目标8",
            外呼下面无目标9 := "中间变量2"."3号梯外呼下面无目标9",
            "1号梯轿内开门按钮" := "输入"."3号梯轿内开门按钮",
            "1号梯轿内关门按钮" := "输入"."3号梯轿内关门按钮",
            上端站1限位 := "输入"."3号梯上端站第1限位",
            下端站1限位 := "输入"."3号梯下端站第1限位",
            "1号梯关门继电器" => "输出"."3号梯关门继电器",
            "1号梯开门继电器" => "输出"."3号梯开门继电器",
            "停梯截断(完成关门）" => "中间变量1"."3号梯停梯截断(置0完成关门）",
            "停梯截断(完成开门）" => "中间变量1"."3号梯停梯截断(置0完成开门）",
            死机 => "中间变量1".死机3);
END_REGION

REGION Network 5: 4
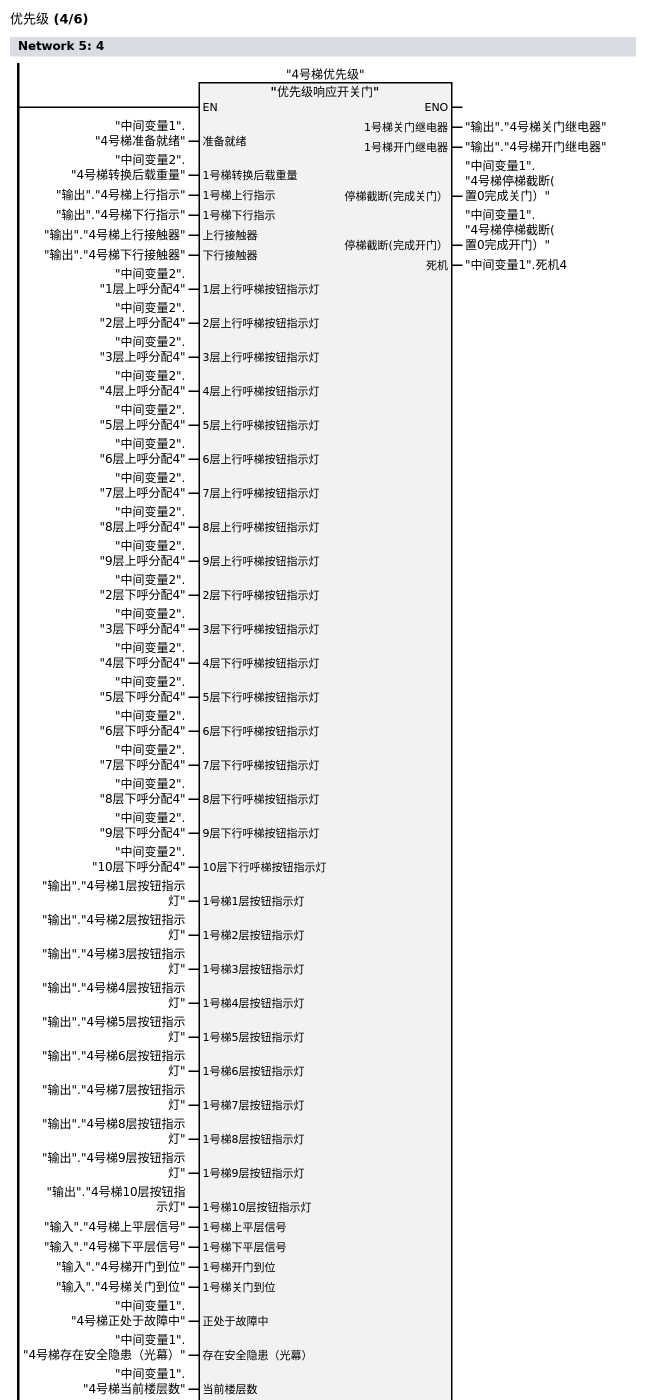
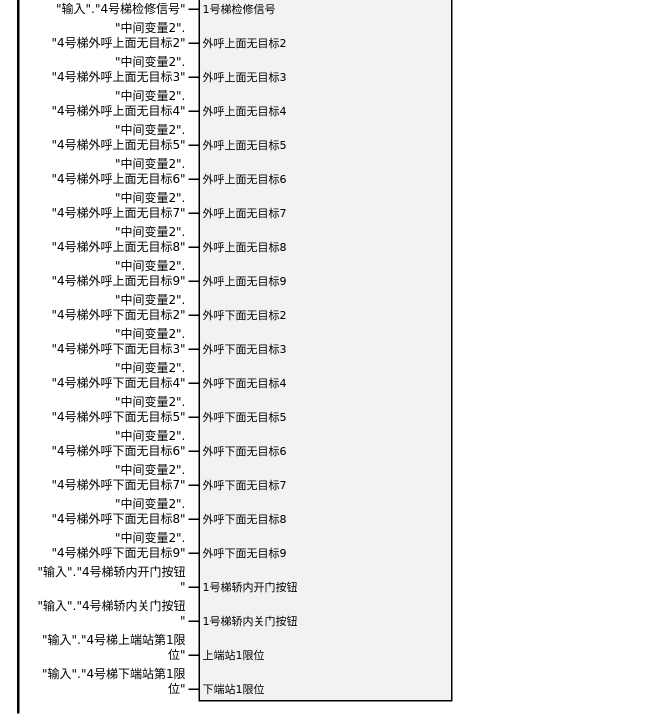
   RUNG wire#powerrail
      "4号梯优先级"(准备就绪 := "中间变量1"."4号梯准备就绪", "1号梯转换后载重量" := "中间变量2"."4号梯转换后载重量", "1号梯上行指示" := "输出"."4号梯上行指示", "1号梯下行指示" := "输出"."4号梯下行指示", 上行接触器 := "输出"."4号梯上行接触器", 下行接触器 := "输出"."4号梯下行接触器", "1层上行呼梯按钮指示灯" := "中间变量2"."1层上呼分配4", "2层上行呼梯按钮指示灯" := "中间变量2"."2层上呼分配4", "3层上行呼梯按钮指示灯" := "中间变量2"."3层上呼分配4", "4层上行呼梯按钮指示灯" := "中间变量2"."4层上呼分配4", "5层上行呼梯按钮指示灯" := "中间变量2"."5层上呼分配4", "6层上行呼梯按钮指示灯" := "中间变量2"."6层上呼分配4", "7层上行呼梯按钮指示灯" := "中间变量2"."7层上呼分配4", "8层上行呼梯按钮指示灯" := "中间变量2"."8层上呼分配4", "9层上行呼梯按钮指示灯" := "中间变量2"."9层上呼分配4", "2层下行呼梯按钮指示灯" := "中间变量2"."2层下呼分配4", "3层下行呼梯按钮指示灯" := "中间变量2"."3层下呼分配4", "4层下行呼梯按钮指示灯" := "中间变量2"."4层下呼分配4", "5层下行呼梯按钮指示灯" := "中间变量2"."5层下呼分配4", "6层下行呼梯按钮指示灯" := "中间变量2"."6层下呼分配4", "7层下行呼梯按钮指示灯" := "中间变量2"."7层下呼分配4", "8层下行呼梯按钮指示灯" := "中间变量2"."8层下呼分配4", "9层下行呼梯按钮指示灯" := "中间变量2"."9层下呼分配4", "10层下行呼梯按钮指示灯" := "中间变量2"."10层下呼分配4", "1号梯1层按钮指示灯" := "输出"."4号梯1层按钮指示灯", "1号梯2层按钮指示灯" := "输出"."4号梯2层按钮指示灯", "1号梯3层按钮指示灯" := "输出"."4号梯3层按钮指示灯", "1号梯4层按钮指示灯" := "输出"."4号梯4层按钮指示灯", "1号梯5层按钮指示灯" := "输出"."4号梯5层按钮指示灯", "1号梯6层按钮指示灯" := "输出"."4号梯6层按钮指示灯", "1号梯7层按钮指示灯" := "输出"."4号梯7层按钮指示灯", "1号梯8层按钮指示灯" := "输出"."4号梯8层按钮指示灯", "1号梯9层按钮指示灯" := "输出"."4号梯9层按钮指示灯", "1号梯10层按钮指示灯" := "输出"."4号梯10层按钮指示灯", "1号梯上平层信号" := "输入"."4号梯上平层信号", "1号梯下平层信号" := "输入"."4号梯下平层信号", "1号梯开门到位" := "输入"."4号梯开门到位", "1号梯关门到位" := "输入"."4号梯关门到位", 正处于故障中 := "中间变量1"."4号梯正处于故障中", "存在安全隐患（光幕）" := "中间变量1"."4号梯存在安全隐患（光幕）", 当前楼层数 := "中间变量1"."4号梯当前楼层数", "1号梯检修信号" := "输入"."4号梯检修信号", 外呼上面无目标2 := "中间变量2"."4号梯外呼上面无目标2", 外呼上面无目标3 := "中间变量2"."4号梯外呼上面无目标3", 外呼上面无目标4 := "中间变量2"."4号梯外呼上面无目标4", 外呼上面无目标5 := "中间变量2"."4号梯外呼上面无目标5", 外呼上面无目标6 := "中间变量2"."4号梯外呼上面无目标6", 外呼上面无目标7 := "中间变量2"."4号梯外呼上面无目标7", 外呼上面无目标8 := "中间变量2"."4号梯外呼上面无目标8", 外呼上面无目标9 := "中间变量2"."4号梯外呼上面无目标9", 外呼下面无目标2 := "中间变量2"."4号梯外呼下面无目标2", 外呼下面无目标3 := "中间变量2"."4号梯外呼下面无目标3", 外呼下面无目标4 := "中间变量2"."4号梯外呼下面无目标4", 外呼下面无目标5 := "中间变量2"."4号梯外呼下面无目标5", 外呼下面无目标6 := "中间变量2"."4号梯外呼下面无目标6", 外呼下面无目标7 := "中间变量2"."4号梯外呼下面无目标7", 外呼下面无目标8 := "中间变量2"."4号梯外呼下面无目标8", 外呼下面无目标9 := "中间变量2"."4号梯外呼下面无目标9", "1号梯轿内开门按钮" := "输入"."4号梯轿内开门按钮", "1号梯轿内关门按钮" := "输入"."4号梯轿内关门按钮", 上端站1限位 := "输入"."4号梯上端站第1限位", 下端站1限位 := "输入"."4号梯下端站第1限位", "1号梯关门继电器" => "输出"."4号梯关门继电器", "1号梯开门继电器" => "输出"."4号梯开门继电器", "停梯截断(完成关门）" => "中间变量1"."4号梯停梯截断(置0完成关门）", "停梯截断(完成开门）" => "中间变量1"."4号梯停梯截断(置0完成开门）", 死机 => "中间变量1".死机4)
   END_RUNG
   // the same network as SCL:
   "4号梯优先级"(准备就绪 := "中间变量1"."4号梯准备就绪",   // "优先级响应开关门"
            "1号梯转换后载重量" := "中间变量2"."4号梯转换后载重量",
            "1号梯上行指示" := "输出"."4号梯上行指示",
            "1号梯下行指示" := "输出"."4号梯下行指示",
            上行接触器 := "输出"."4号梯上行接触器",
            下行接触器 := "输出"."4号梯下行接触器",
            "1层上行呼梯按钮指示灯" := "中间变量2"."1层上呼分配4",
            "2层上行呼梯按钮指示灯" := "中间变量2"."2层上呼分配4",
            "3层上行呼梯按钮指示灯" := "中间变量2"."3层上呼分配4",
            "4层上行呼梯按钮指示灯" := "中间变量2"."4层上呼分配4",
            "5层上行呼梯按钮指示灯" := "中间变量2"."5层上呼分配4",
            "6层上行呼梯按钮指示灯" := "中间变量2"."6层上呼分配4",
            "7层上行呼梯按钮指示灯" := "中间变量2"."7层上呼分配4",
            "8层上行呼梯按钮指示灯" := "中间变量2"."8层上呼分配4",
            "9层上行呼梯按钮指示灯" := "中间变量2"."9层上呼分配4",
            "2层下行呼梯按钮指示灯" := "中间变量2"."2层下呼分配4",
            "3层下行呼梯按钮指示灯" := "中间变量2"."3层下呼分配4",
            "4层下行呼梯按钮指示灯" := "中间变量2"."4层下呼分配4",
            "5层下行呼梯按钮指示灯" := "中间变量2"."5层下呼分配4",
            "6层下行呼梯按钮指示灯" := "中间变量2"."6层下呼分配4",
            "7层下行呼梯按钮指示灯" := "中间变量2"."7层下呼分配4",
            "8层下行呼梯按钮指示灯" := "中间变量2"."8层下呼分配4",
            "9层下行呼梯按钮指示灯" := "中间变量2"."9层下呼分配4",
            "10层下行呼梯按钮指示灯" := "中间变量2"."10层下呼分配4",
            "1号梯1层按钮指示灯" := "输出"."4号梯1层按钮指示灯",
            "1号梯2层按钮指示灯" := "输出"."4号梯2层按钮指示灯",
            "1号梯3层按钮指示灯" := "输出"."4号梯3层按钮指示灯",
            "1号梯4层按钮指示灯" := "输出"."4号梯4层按钮指示灯",
            "1号梯5层按钮指示灯" := "输出"."4号梯5层按钮指示灯",
            "1号梯6层按钮指示灯" := "输出"."4号梯6层按钮指示灯",
            "1号梯7层按钮指示灯" := "输出"."4号梯7层按钮指示灯",
            "1号梯8层按钮指示灯" := "输出"."4号梯8层按钮指示灯",
            "1号梯9层按钮指示灯" := "输出"."4号梯9层按钮指示灯",
            "1号梯10层按钮指示灯" := "输出"."4号梯10层按钮指示灯",
            "1号梯上平层信号" := "输入"."4号梯上平层信号",
            "1号梯下平层信号" := "输入"."4号梯下平层信号",
            "1号梯开门到位" := "输入"."4号梯开门到位",
            "1号梯关门到位" := "输入"."4号梯关门到位",
            正处于故障中 := "中间变量1"."4号梯正处于故障中",
            "存在安全隐患（光幕）" := "中间变量1"."4号梯存在安全隐患（光幕）",
            当前楼层数 := "中间变量1"."4号梯当前楼层数",
            "1号梯检修信号" := "输入"."4号梯检修信号",
            外呼上面无目标2 := "中间变量2"."4号梯外呼上面无目标2",
            外呼上面无目标3 := "中间变量2"."4号梯外呼上面无目标3",
            外呼上面无目标4 := "中间变量2"."4号梯外呼上面无目标4",
            外呼上面无目标5 := "中间变量2"."4号梯外呼上面无目标5",
            外呼上面无目标6 := "中间变量2"."4号梯外呼上面无目标6",
            外呼上面无目标7 := "中间变量2"."4号梯外呼上面无目标7",
            外呼上面无目标8 := "中间变量2"."4号梯外呼上面无目标8",
            外呼上面无目标9 := "中间变量2"."4号梯外呼上面无目标9",
            外呼下面无目标2 := "中间变量2"."4号梯外呼下面无目标2",
            外呼下面无目标3 := "中间变量2"."4号梯外呼下面无目标3",
            外呼下面无目标4 := "中间变量2"."4号梯外呼下面无目标4",
            外呼下面无目标5 := "中间变量2"."4号梯外呼下面无目标5",
            外呼下面无目标6 := "中间变量2"."4号梯外呼下面无目标6",
            外呼下面无目标7 := "中间变量2"."4号梯外呼下面无目标7",
            外呼下面无目标8 := "中间变量2"."4号梯外呼下面无目标8",
            外呼下面无目标9 := "中间变量2"."4号梯外呼下面无目标9",
            "1号梯轿内开门按钮" := "输入"."4号梯轿内开门按钮",
            "1号梯轿内关门按钮" := "输入"."4号梯轿内关门按钮",
            上端站1限位 := "输入"."4号梯上端站第1限位",
            下端站1限位 := "输入"."4号梯下端站第1限位",
            "1号梯关门继电器" => "输出"."4号梯关门继电器",
            "1号梯开门继电器" => "输出"."4号梯开门继电器",
            "停梯截断(完成关门）" => "中间变量1"."4号梯停梯截断(置0完成关门）",
            "停梯截断(完成开门）" => "中间变量1"."4号梯停梯截断(置0完成开门）",
            死机 => "中间变量1".死机4);
END_REGION

REGION Network 6: 5
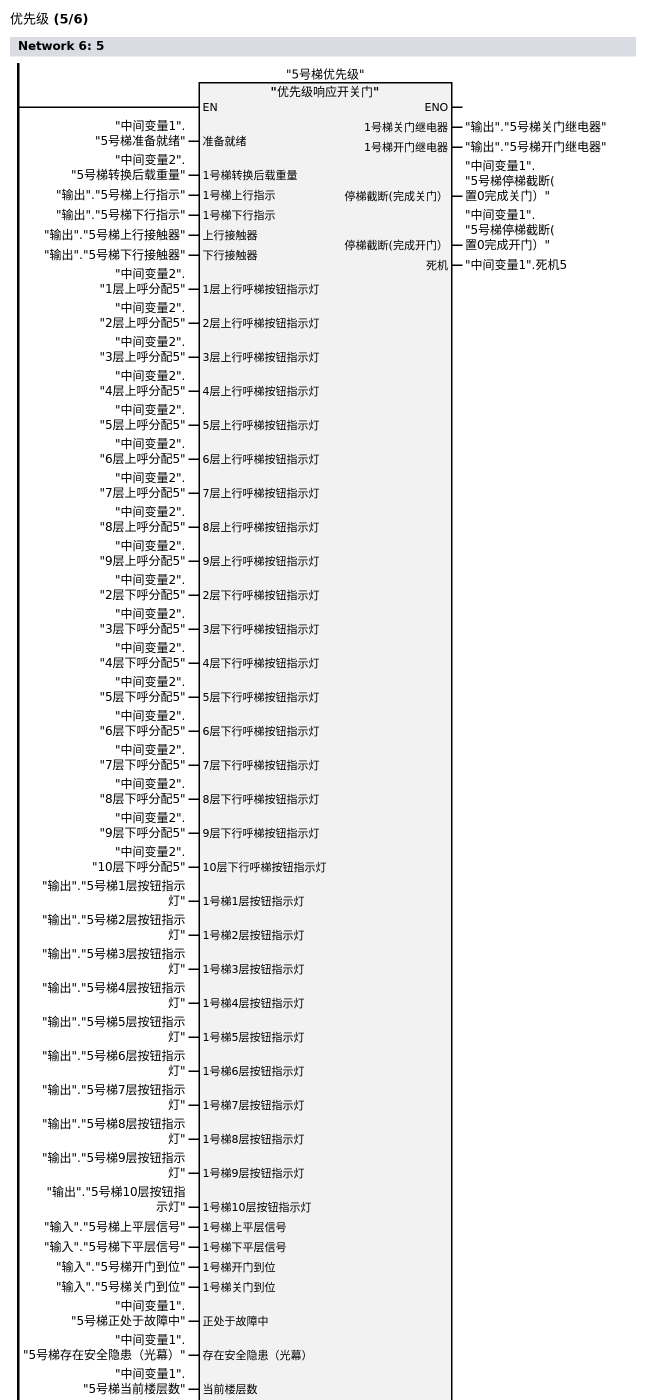
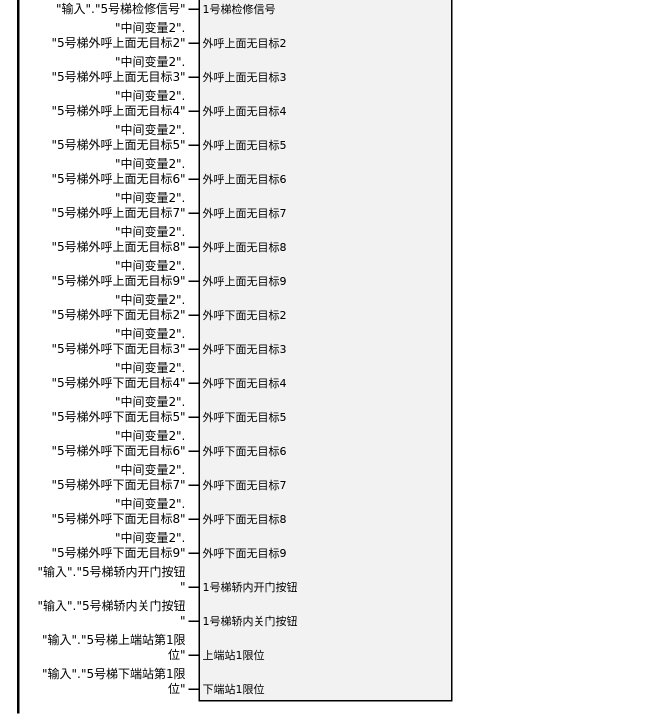
   RUNG wire#powerrail
      "5号梯优先级"(准备就绪 := "中间变量1"."5号梯准备就绪", "1号梯转换后载重量" := "中间变量2"."5号梯转换后载重量", "1号梯上行指示" := "输出"."5号梯上行指示", "1号梯下行指示" := "输出"."5号梯下行指示", 上行接触器 := "输出"."5号梯上行接触器", 下行接触器 := "输出"."5号梯下行接触器", "1层上行呼梯按钮指示灯" := "中间变量2"."1层上呼分配5", "2层上行呼梯按钮指示灯" := "中间变量2"."2层上呼分配5", "3层上行呼梯按钮指示灯" := "中间变量2"."3层上呼分配5", "4层上行呼梯按钮指示灯" := "中间变量2"."4层上呼分配5", "5层上行呼梯按钮指示灯" := "中间变量2"."5层上呼分配5", "6层上行呼梯按钮指示灯" := "中间变量2"."6层上呼分配5", "7层上行呼梯按钮指示灯" := "中间变量2"."7层上呼分配5", "8层上行呼梯按钮指示灯" := "中间变量2"."8层上呼分配5", "9层上行呼梯按钮指示灯" := "中间变量2"."9层上呼分配5", "2层下行呼梯按钮指示灯" := "中间变量2"."2层下呼分配5", "3层下行呼梯按钮指示灯" := "中间变量2"."3层下呼分配5", "4层下行呼梯按钮指示灯" := "中间变量2"."4层下呼分配5", "5层下行呼梯按钮指示灯" := "中间变量2"."5层下呼分配5", "6层下行呼梯按钮指示灯" := "中间变量2"."6层下呼分配5", "7层下行呼梯按钮指示灯" := "中间变量2"."7层下呼分配5", "8层下行呼梯按钮指示灯" := "中间变量2"."8层下呼分配5", "9层下行呼梯按钮指示灯" := "中间变量2"."9层下呼分配5", "10层下行呼梯按钮指示灯" := "中间变量2"."10层下呼分配5", "1号梯1层按钮指示灯" := "输出"."5号梯1层按钮指示灯", "1号梯2层按钮指示灯" := "输出"."5号梯2层按钮指示灯", "1号梯3层按钮指示灯" := "输出"."5号梯3层按钮指示灯", "1号梯4层按钮指示灯" := "输出"."5号梯4层按钮指示灯", "1号梯5层按钮指示灯" := "输出"."5号梯5层按钮指示灯", "1号梯6层按钮指示灯" := "输出"."5号梯6层按钮指示灯", "1号梯7层按钮指示灯" := "输出"."5号梯7层按钮指示灯", "1号梯8层按钮指示灯" := "输出"."5号梯8层按钮指示灯", "1号梯9层按钮指示灯" := "输出"."5号梯9层按钮指示灯", "1号梯10层按钮指示灯" := "输出"."5号梯10层按钮指示灯", "1号梯上平层信号" := "输入"."5号梯上平层信号", "1号梯下平层信号" := "输入"."5号梯下平层信号", "1号梯开门到位" := "输入"."5号梯开门到位", "1号梯关门到位" := "输入"."5号梯关门到位", 正处于故障中 := "中间变量1"."5号梯正处于故障中", "存在安全隐患（光幕）" := "中间变量1"."5号梯存在安全隐患（光幕）", 当前楼层数 := "中间变量1"."5号梯当前楼层数", "1号梯检修信号" := "输入"."5号梯检修信号", 外呼上面无目标2 := "中间变量2"."5号梯外呼上面无目标2", 外呼上面无目标3 := "中间变量2"."5号梯外呼上面无目标3", 外呼上面无目标4 := "中间变量2"."5号梯外呼上面无目标4", 外呼上面无目标5 := "中间变量2"."5号梯外呼上面无目标5", 外呼上面无目标6 := "中间变量2"."5号梯外呼上面无目标6", 外呼上面无目标7 := "中间变量2"."5号梯外呼上面无目标7", 外呼上面无目标8 := "中间变量2"."5号梯外呼上面无目标8", 外呼上面无目标9 := "中间变量2"."5号梯外呼上面无目标9", 外呼下面无目标2 := "中间变量2"."5号梯外呼下面无目标2", 外呼下面无目标3 := "中间变量2"."5号梯外呼下面无目标3", 外呼下面无目标4 := "中间变量2"."5号梯外呼下面无目标4", 外呼下面无目标5 := "中间变量2"."5号梯外呼下面无目标5", 外呼下面无目标6 := "中间变量2"."5号梯外呼下面无目标6", 外呼下面无目标7 := "中间变量2"."5号梯外呼下面无目标7", 外呼下面无目标8 := "中间变量2"."5号梯外呼下面无目标8", 外呼下面无目标9 := "中间变量2"."5号梯外呼下面无目标9", "1号梯轿内开门按钮" := "输入"."5号梯轿内开门按钮", "1号梯轿内关门按钮" := "输入"."5号梯轿内关门按钮", 上端站1限位 := "输入"."5号梯上端站第1限位", 下端站1限位 := "输入"."5号梯下端站第1限位", "1号梯关门继电器" => "输出"."5号梯关门继电器", "1号梯开门继电器" => "输出"."5号梯开门继电器", "停梯截断(完成关门）" => "中间变量1"."5号梯停梯截断(置0完成关门）", "停梯截断(完成开门）" => "中间变量1"."5号梯停梯截断(置0完成开门）", 死机 => "中间变量1".死机5)
   END_RUNG
   // the same network as SCL:
   "5号梯优先级"(准备就绪 := "中间变量1"."5号梯准备就绪",   // "优先级响应开关门"
            "1号梯转换后载重量" := "中间变量2"."5号梯转换后载重量",
            "1号梯上行指示" := "输出"."5号梯上行指示",
            "1号梯下行指示" := "输出"."5号梯下行指示",
            上行接触器 := "输出"."5号梯上行接触器",
            下行接触器 := "输出"."5号梯下行接触器",
            "1层上行呼梯按钮指示灯" := "中间变量2"."1层上呼分配5",
            "2层上行呼梯按钮指示灯" := "中间变量2"."2层上呼分配5",
            "3层上行呼梯按钮指示灯" := "中间变量2"."3层上呼分配5",
            "4层上行呼梯按钮指示灯" := "中间变量2"."4层上呼分配5",
            "5层上行呼梯按钮指示灯" := "中间变量2"."5层上呼分配5",
            "6层上行呼梯按钮指示灯" := "中间变量2"."6层上呼分配5",
            "7层上行呼梯按钮指示灯" := "中间变量2"."7层上呼分配5",
            "8层上行呼梯按钮指示灯" := "中间变量2"."8层上呼分配5",
            "9层上行呼梯按钮指示灯" := "中间变量2"."9层上呼分配5",
            "2层下行呼梯按钮指示灯" := "中间变量2"."2层下呼分配5",
            "3层下行呼梯按钮指示灯" := "中间变量2"."3层下呼分配5",
            "4层下行呼梯按钮指示灯" := "中间变量2"."4层下呼分配5",
            "5层下行呼梯按钮指示灯" := "中间变量2"."5层下呼分配5",
            "6层下行呼梯按钮指示灯" := "中间变量2"."6层下呼分配5",
            "7层下行呼梯按钮指示灯" := "中间变量2"."7层下呼分配5",
            "8层下行呼梯按钮指示灯" := "中间变量2"."8层下呼分配5",
            "9层下行呼梯按钮指示灯" := "中间变量2"."9层下呼分配5",
            "10层下行呼梯按钮指示灯" := "中间变量2"."10层下呼分配5",
            "1号梯1层按钮指示灯" := "输出"."5号梯1层按钮指示灯",
            "1号梯2层按钮指示灯" := "输出"."5号梯2层按钮指示灯",
            "1号梯3层按钮指示灯" := "输出"."5号梯3层按钮指示灯",
            "1号梯4层按钮指示灯" := "输出"."5号梯4层按钮指示灯",
            "1号梯5层按钮指示灯" := "输出"."5号梯5层按钮指示灯",
            "1号梯6层按钮指示灯" := "输出"."5号梯6层按钮指示灯",
            "1号梯7层按钮指示灯" := "输出"."5号梯7层按钮指示灯",
            "1号梯8层按钮指示灯" := "输出"."5号梯8层按钮指示灯",
            "1号梯9层按钮指示灯" := "输出"."5号梯9层按钮指示灯",
            "1号梯10层按钮指示灯" := "输出"."5号梯10层按钮指示灯",
            "1号梯上平层信号" := "输入"."5号梯上平层信号",
            "1号梯下平层信号" := "输入"."5号梯下平层信号",
            "1号梯开门到位" := "输入"."5号梯开门到位",
            "1号梯关门到位" := "输入"."5号梯关门到位",
            正处于故障中 := "中间变量1"."5号梯正处于故障中",
            "存在安全隐患（光幕）" := "中间变量1"."5号梯存在安全隐患（光幕）",
            当前楼层数 := "中间变量1"."5号梯当前楼层数",
            "1号梯检修信号" := "输入"."5号梯检修信号",
            外呼上面无目标2 := "中间变量2"."5号梯外呼上面无目标2",
            外呼上面无目标3 := "中间变量2"."5号梯外呼上面无目标3",
            外呼上面无目标4 := "中间变量2"."5号梯外呼上面无目标4",
            外呼上面无目标5 := "中间变量2"."5号梯外呼上面无目标5",
            外呼上面无目标6 := "中间变量2"."5号梯外呼上面无目标6",
            外呼上面无目标7 := "中间变量2"."5号梯外呼上面无目标7",
            外呼上面无目标8 := "中间变量2"."5号梯外呼上面无目标8",
            外呼上面无目标9 := "中间变量2"."5号梯外呼上面无目标9",
            外呼下面无目标2 := "中间变量2"."5号梯外呼下面无目标2",
            外呼下面无目标3 := "中间变量2"."5号梯外呼下面无目标3",
            外呼下面无目标4 := "中间变量2"."5号梯外呼下面无目标4",
            外呼下面无目标5 := "中间变量2"."5号梯外呼下面无目标5",
            外呼下面无目标6 := "中间变量2"."5号梯外呼下面无目标6",
            外呼下面无目标7 := "中间变量2"."5号梯外呼下面无目标7",
            外呼下面无目标8 := "中间变量2"."5号梯外呼下面无目标8",
            外呼下面无目标9 := "中间变量2"."5号梯外呼下面无目标9",
            "1号梯轿内开门按钮" := "输入"."5号梯轿内开门按钮",
            "1号梯轿内关门按钮" := "输入"."5号梯轿内关门按钮",
            上端站1限位 := "输入"."5号梯上端站第1限位",
            下端站1限位 := "输入"."5号梯下端站第1限位",
            "1号梯关门继电器" => "输出"."5号梯关门继电器",
            "1号梯开门继电器" => "输出"."5号梯开门继电器",
            "停梯截断(完成关门）" => "中间变量1"."5号梯停梯截断(置0完成关门）",
            "停梯截断(完成开门）" => "中间变量1"."5号梯停梯截断(置0完成开门）",
            死机 => "中间变量1".死机5);
END_REGION

REGION Network 7: 6
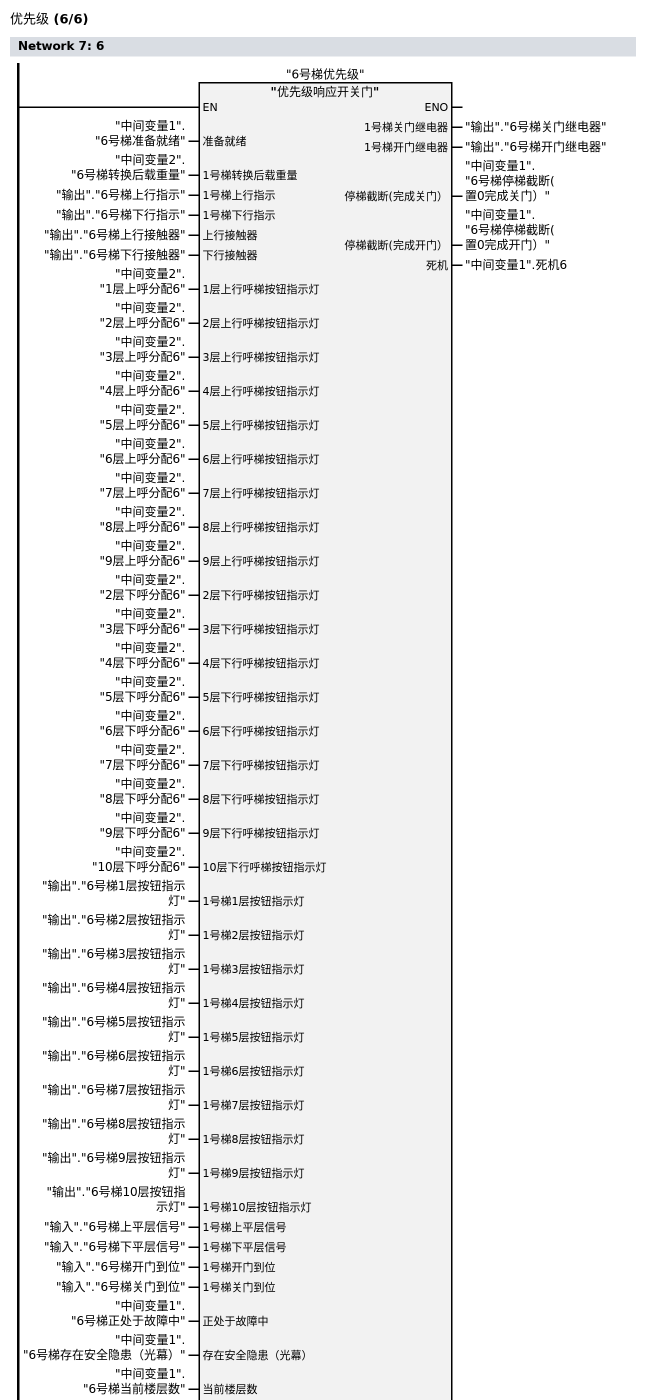
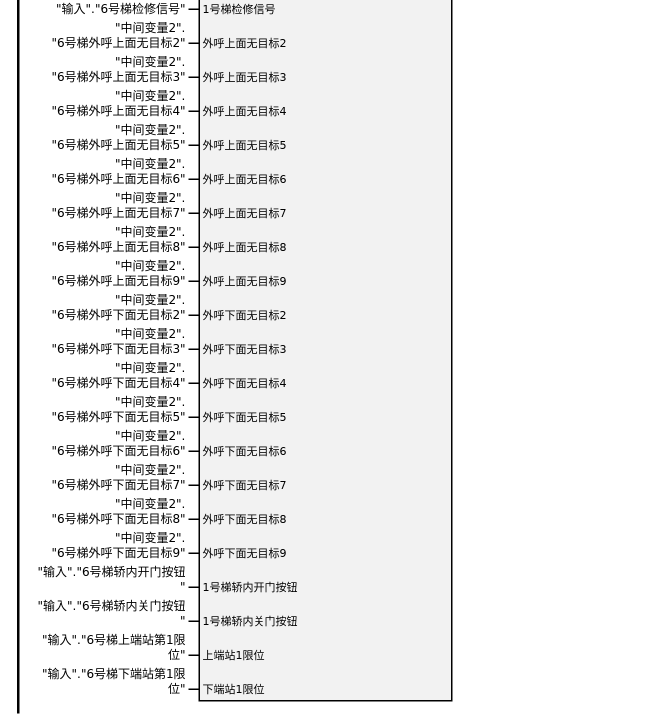
   RUNG wire#powerrail
      "6号梯优先级"(准备就绪 := "中间变量1"."6号梯准备就绪", "1号梯转换后载重量" := "中间变量2"."6号梯转换后载重量", "1号梯上行指示" := "输出"."6号梯上行指示", "1号梯下行指示" := "输出"."6号梯下行指示", 上行接触器 := "输出"."6号梯上行接触器", 下行接触器 := "输出"."6号梯下行接触器", "1层上行呼梯按钮指示灯" := "中间变量2"."1层上呼分配6", "2层上行呼梯按钮指示灯" := "中间变量2"."2层上呼分配6", "3层上行呼梯按钮指示灯" := "中间变量2"."3层上呼分配6", "4层上行呼梯按钮指示灯" := "中间变量2"."4层上呼分配6", "5层上行呼梯按钮指示灯" := "中间变量2"."5层上呼分配6", "6层上行呼梯按钮指示灯" := "中间变量2"."6层上呼分配6", "7层上行呼梯按钮指示灯" := "中间变量2"."7层上呼分配6", "8层上行呼梯按钮指示灯" := "中间变量2"."8层上呼分配6", "9层上行呼梯按钮指示灯" := "中间变量2"."9层上呼分配6", "2层下行呼梯按钮指示灯" := "中间变量2"."2层下呼分配6", "3层下行呼梯按钮指示灯" := "中间变量2"."3层下呼分配6", "4层下行呼梯按钮指示灯" := "中间变量2"."4层下呼分配6", "5层下行呼梯按钮指示灯" := "中间变量2"."5层下呼分配6", "6层下行呼梯按钮指示灯" := "中间变量2"."6层下呼分配6", "7层下行呼梯按钮指示灯" := "中间变量2"."7层下呼分配6", "8层下行呼梯按钮指示灯" := "中间变量2"."8层下呼分配6", "9层下行呼梯按钮指示灯" := "中间变量2"."9层下呼分配6", "10层下行呼梯按钮指示灯" := "中间变量2"."10层下呼分配6", "1号梯1层按钮指示灯" := "输出"."6号梯1层按钮指示灯", "1号梯2层按钮指示灯" := "输出"."6号梯2层按钮指示灯", "1号梯3层按钮指示灯" := "输出"."6号梯3层按钮指示灯", "1号梯4层按钮指示灯" := "输出"."6号梯4层按钮指示灯", "1号梯5层按钮指示灯" := "输出"."6号梯5层按钮指示灯", "1号梯6层按钮指示灯" := "输出"."6号梯6层按钮指示灯", "1号梯7层按钮指示灯" := "输出"."6号梯7层按钮指示灯", "1号梯8层按钮指示灯" := "输出"."6号梯8层按钮指示灯", "1号梯9层按钮指示灯" := "输出"."6号梯9层按钮指示灯", "1号梯10层按钮指示灯" := "输出"."6号梯10层按钮指示灯", "1号梯上平层信号" := "输入"."6号梯上平层信号", "1号梯下平层信号" := "输入"."6号梯下平层信号", "1号梯开门到位" := "输入"."6号梯开门到位", "1号梯关门到位" := "输入"."6号梯关门到位", 正处于故障中 := "中间变量1"."6号梯正处于故障中", "存在安全隐患（光幕）" := "中间变量1"."6号梯存在安全隐患（光幕）", 当前楼层数 := "中间变量1"."6号梯当前楼层数", "1号梯检修信号" := "输入"."6号梯检修信号", 外呼上面无目标2 := "中间变量2"."6号梯外呼上面无目标2", 外呼上面无目标3 := "中间变量2"."6号梯外呼上面无目标3", 外呼上面无目标4 := "中间变量2"."6号梯外呼上面无目标4", 外呼上面无目标5 := "中间变量2"."6号梯外呼上面无目标5", 外呼上面无目标6 := "中间变量2"."6号梯外呼上面无目标6", 外呼上面无目标7 := "中间变量2"."6号梯外呼上面无目标7", 外呼上面无目标8 := "中间变量2"."6号梯外呼上面无目标8", 外呼上面无目标9 := "中间变量2"."6号梯外呼上面无目标9", 外呼下面无目标2 := "中间变量2"."6号梯外呼下面无目标2", 外呼下面无目标3 := "中间变量2"."6号梯外呼下面无目标3", 外呼下面无目标4 := "中间变量2"."6号梯外呼下面无目标4", 外呼下面无目标5 := "中间变量2"."6号梯外呼下面无目标5", 外呼下面无目标6 := "中间变量2"."6号梯外呼下面无目标6", 外呼下面无目标7 := "中间变量2"."6号梯外呼下面无目标7", 外呼下面无目标8 := "中间变量2"."6号梯外呼下面无目标8", 外呼下面无目标9 := "中间变量2"."6号梯外呼下面无目标9", "1号梯轿内开门按钮" := "输入"."6号梯轿内开门按钮", "1号梯轿内关门按钮" := "输入"."6号梯轿内关门按钮", 上端站1限位 := "输入"."6号梯上端站第1限位", 下端站1限位 := "输入"."6号梯下端站第1限位", "1号梯关门继电器" => "输出"."6号梯关门继电器", "1号梯开门继电器" => "输出"."6号梯开门继电器", "停梯截断(完成关门）" => "中间变量1"."6号梯停梯截断(置0完成关门）", "停梯截断(完成开门）" => "中间变量1"."6号梯停梯截断(置0完成开门）", 死机 => "中间变量1".死机6)
   END_RUNG
   // the same network as SCL:
   "6号梯优先级"(准备就绪 := "中间变量1"."6号梯准备就绪",   // "优先级响应开关门"
            "1号梯转换后载重量" := "中间变量2"."6号梯转换后载重量",
            "1号梯上行指示" := "输出"."6号梯上行指示",
            "1号梯下行指示" := "输出"."6号梯下行指示",
            上行接触器 := "输出"."6号梯上行接触器",
            下行接触器 := "输出"."6号梯下行接触器",
            "1层上行呼梯按钮指示灯" := "中间变量2"."1层上呼分配6",
            "2层上行呼梯按钮指示灯" := "中间变量2"."2层上呼分配6",
            "3层上行呼梯按钮指示灯" := "中间变量2"."3层上呼分配6",
            "4层上行呼梯按钮指示灯" := "中间变量2"."4层上呼分配6",
            "5层上行呼梯按钮指示灯" := "中间变量2"."5层上呼分配6",
            "6层上行呼梯按钮指示灯" := "中间变量2"."6层上呼分配6",
            "7层上行呼梯按钮指示灯" := "中间变量2"."7层上呼分配6",
            "8层上行呼梯按钮指示灯" := "中间变量2"."8层上呼分配6",
            "9层上行呼梯按钮指示灯" := "中间变量2"."9层上呼分配6",
            "2层下行呼梯按钮指示灯" := "中间变量2"."2层下呼分配6",
            "3层下行呼梯按钮指示灯" := "中间变量2"."3层下呼分配6",
            "4层下行呼梯按钮指示灯" := "中间变量2"."4层下呼分配6",
            "5层下行呼梯按钮指示灯" := "中间变量2"."5层下呼分配6",
            "6层下行呼梯按钮指示灯" := "中间变量2"."6层下呼分配6",
            "7层下行呼梯按钮指示灯" := "中间变量2"."7层下呼分配6",
            "8层下行呼梯按钮指示灯" := "中间变量2"."8层下呼分配6",
            "9层下行呼梯按钮指示灯" := "中间变量2"."9层下呼分配6",
            "10层下行呼梯按钮指示灯" := "中间变量2"."10层下呼分配6",
            "1号梯1层按钮指示灯" := "输出"."6号梯1层按钮指示灯",
            "1号梯2层按钮指示灯" := "输出"."6号梯2层按钮指示灯",
            "1号梯3层按钮指示灯" := "输出"."6号梯3层按钮指示灯",
            "1号梯4层按钮指示灯" := "输出"."6号梯4层按钮指示灯",
            "1号梯5层按钮指示灯" := "输出"."6号梯5层按钮指示灯",
            "1号梯6层按钮指示灯" := "输出"."6号梯6层按钮指示灯",
            "1号梯7层按钮指示灯" := "输出"."6号梯7层按钮指示灯",
            "1号梯8层按钮指示灯" := "输出"."6号梯8层按钮指示灯",
            "1号梯9层按钮指示灯" := "输出"."6号梯9层按钮指示灯",
            "1号梯10层按钮指示灯" := "输出"."6号梯10层按钮指示灯",
            "1号梯上平层信号" := "输入"."6号梯上平层信号",
            "1号梯下平层信号" := "输入"."6号梯下平层信号",
            "1号梯开门到位" := "输入"."6号梯开门到位",
            "1号梯关门到位" := "输入"."6号梯关门到位",
            正处于故障中 := "中间变量1"."6号梯正处于故障中",
            "存在安全隐患（光幕）" := "中间变量1"."6号梯存在安全隐患（光幕）",
            当前楼层数 := "中间变量1"."6号梯当前楼层数",
            "1号梯检修信号" := "输入"."6号梯检修信号",
            外呼上面无目标2 := "中间变量2"."6号梯外呼上面无目标2",
            外呼上面无目标3 := "中间变量2"."6号梯外呼上面无目标3",
            外呼上面无目标4 := "中间变量2"."6号梯外呼上面无目标4",
            外呼上面无目标5 := "中间变量2"."6号梯外呼上面无目标5",
            外呼上面无目标6 := "中间变量2"."6号梯外呼上面无目标6",
            外呼上面无目标7 := "中间变量2"."6号梯外呼上面无目标7",
            外呼上面无目标8 := "中间变量2"."6号梯外呼上面无目标8",
            外呼上面无目标9 := "中间变量2"."6号梯外呼上面无目标9",
            外呼下面无目标2 := "中间变量2"."6号梯外呼下面无目标2",
            外呼下面无目标3 := "中间变量2"."6号梯外呼下面无目标3",
            外呼下面无目标4 := "中间变量2"."6号梯外呼下面无目标4",
            外呼下面无目标5 := "中间变量2"."6号梯外呼下面无目标5",
            外呼下面无目标6 := "中间变量2"."6号梯外呼下面无目标6",
            外呼下面无目标7 := "中间变量2"."6号梯外呼下面无目标7",
            外呼下面无目标8 := "中间变量2"."6号梯外呼下面无目标8",
            外呼下面无目标9 := "中间变量2"."6号梯外呼下面无目标9",
            "1号梯轿内开门按钮" := "输入"."6号梯轿内开门按钮",
            "1号梯轿内关门按钮" := "输入"."6号梯轿内关门按钮",
            上端站1限位 := "输入"."6号梯上端站第1限位",
            下端站1限位 := "输入"."6号梯下端站第1限位",
            "1号梯关门继电器" => "输出"."6号梯关门继电器",
            "1号梯开门继电器" => "输出"."6号梯开门继电器",
            "停梯截断(完成关门）" => "中间变量1"."6号梯停梯截断(置0完成关门）",
            "停梯截断(完成开门）" => "中间变量1"."6号梯停梯截断(置0完成开门）",
            死机 => "中间变量1".死机6);
END_REGION
END_FUNCTION

FUNCTION "指示灯汇总" : Void   // FC11, LAD
{ S7_Optimized_Access := 'TRUE' }
VERSION : 0.1
BEGIN

REGION Network 1: 1号梯指示灯
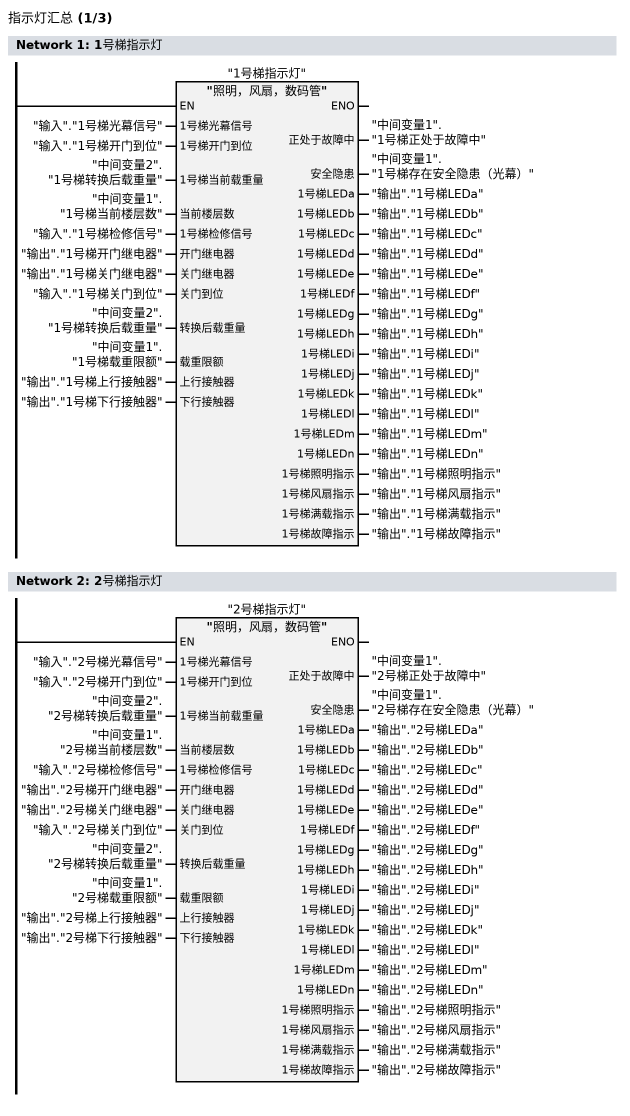
   RUNG wire#powerrail
      "1号梯指示灯"("1号梯光幕信号" := "输入"."1号梯光幕信号", "1号梯开门到位" := "输入"."1号梯开门到位", "1号梯当前载重量" := "中间变量2"."1号梯转换后载重量", 当前楼层数 := "中间变量1"."1号梯当前楼层数", "1号梯检修信号" := "输入"."1号梯检修信号", 开门继电器 := "输出"."1号梯开门继电器", 关门继电器 := "输出"."1号梯关门继电器", 关门到位 := "输入"."1号梯关门到位", 转换后载重量 := "中间变量2"."1号梯转换后载重量", 载重限额 := "中间变量1"."1号梯载重限额", 上行接触器 := "输出"."1号梯上行接触器", 下行接触器 := "输出"."1号梯下行接触器", 正处于故障中 => "中间变量1"."1号梯正处于故障中", 安全隐患 => "中间变量1"."1号梯存在安全隐患（光幕）", "1号梯LEDa" => "输出"."1号梯LEDa", "1号梯LEDb" => "输出"."1号梯LEDb", "1号梯LEDc" => "输出"."1号梯LEDc", "1号梯LEDd" => "输出"."1号梯LEDd", "1号梯LEDe" => "输出"."1号梯LEDe", "1号梯LEDf" => "输出"."1号梯LEDf", "1号梯LEDg" => "输出"."1号梯LEDg", "1号梯LEDh" => "输出"."1号梯LEDh", "1号梯LEDi" => "输出"."1号梯LEDi", "1号梯LEDj" => "输出"."1号梯LEDj", "1号梯LEDk" => "输出"."1号梯LEDk", "1号梯LEDl" => "输出"."1号梯LEDl", "1号梯LEDm" => "输出"."1号梯LEDm", "1号梯LEDn" => "输出"."1号梯LEDn", "1号梯照明指示" => "输出"."1号梯照明指示", "1号梯风扇指示" => "输出"."1号梯风扇指示", "1号梯满载指示" => "输出"."1号梯满载指示", "1号梯故障指示" => "输出"."1号梯故障指示")
   END_RUNG
   // the same network as SCL:
   "1号梯指示灯"("1号梯光幕信号" := "输入"."1号梯光幕信号",   // "照明，风扇，数码管"
            "1号梯开门到位" := "输入"."1号梯开门到位",
            "1号梯当前载重量" := "中间变量2"."1号梯转换后载重量",
            当前楼层数 := "中间变量1"."1号梯当前楼层数",
            "1号梯检修信号" := "输入"."1号梯检修信号",
            开门继电器 := "输出"."1号梯开门继电器",
            关门继电器 := "输出"."1号梯关门继电器",
            关门到位 := "输入"."1号梯关门到位",
            转换后载重量 := "中间变量2"."1号梯转换后载重量",
            载重限额 := "中间变量1"."1号梯载重限额",
            上行接触器 := "输出"."1号梯上行接触器",
            下行接触器 := "输出"."1号梯下行接触器",
            正处于故障中 => "中间变量1"."1号梯正处于故障中",
            安全隐患 => "中间变量1"."1号梯存在安全隐患（光幕）",
            "1号梯LEDa" => "输出"."1号梯LEDa",
            "1号梯LEDb" => "输出"."1号梯LEDb",
            "1号梯LEDc" => "输出"."1号梯LEDc",
            "1号梯LEDd" => "输出"."1号梯LEDd",
            "1号梯LEDe" => "输出"."1号梯LEDe",
            "1号梯LEDf" => "输出"."1号梯LEDf",
            "1号梯LEDg" => "输出"."1号梯LEDg",
            "1号梯LEDh" => "输出"."1号梯LEDh",
            "1号梯LEDi" => "输出"."1号梯LEDi",
            "1号梯LEDj" => "输出"."1号梯LEDj",
            "1号梯LEDk" => "输出"."1号梯LEDk",
            "1号梯LEDl" => "输出"."1号梯LEDl",
            "1号梯LEDm" => "输出"."1号梯LEDm",
            "1号梯LEDn" => "输出"."1号梯LEDn",
            "1号梯照明指示" => "输出"."1号梯照明指示",
            "1号梯风扇指示" => "输出"."1号梯风扇指示",
            "1号梯满载指示" => "输出"."1号梯满载指示",
            "1号梯故障指示" => "输出"."1号梯故障指示");
END_REGION

REGION Network 2: 2号梯指示灯
   RUNG wire#powerrail
      "2号梯指示灯"("1号梯光幕信号" := "输入"."2号梯光幕信号", "1号梯开门到位" := "输入"."2号梯开门到位", "1号梯当前载重量" := "中间变量2"."2号梯转换后载重量", 当前楼层数 := "中间变量1"."2号梯当前楼层数", "1号梯检修信号" := "输入"."2号梯检修信号", 开门继电器 := "输出"."2号梯开门继电器", 关门继电器 := "输出"."2号梯关门继电器", 关门到位 := "输入"."2号梯关门到位", 转换后载重量 := "中间变量2"."2号梯转换后载重量", 载重限额 := "中间变量1"."2号梯载重限额", 上行接触器 := "输出"."2号梯上行接触器", 下行接触器 := "输出"."2号梯下行接触器", 正处于故障中 => "中间变量1"."2号梯正处于故障中", 安全隐患 => "中间变量1"."2号梯存在安全隐患（光幕）", "1号梯LEDa" => "输出"."2号梯LEDa", "1号梯LEDb" => "输出"."2号梯LEDb", "1号梯LEDc" => "输出"."2号梯LEDc", "1号梯LEDd" => "输出"."2号梯LEDd", "1号梯LEDe" => "输出"."2号梯LEDe", "1号梯LEDf" => "输出"."2号梯LEDf", "1号梯LEDg" => "输出"."2号梯LEDg", "1号梯LEDh" => "输出"."2号梯LEDh", "1号梯LEDi" => "输出"."2号梯LEDi", "1号梯LEDj" => "输出"."2号梯LEDj", "1号梯LEDk" => "输出"."2号梯LEDk", "1号梯LEDl" => "输出"."2号梯LEDl", "1号梯LEDm" => "输出"."2号梯LEDm", "1号梯LEDn" => "输出"."2号梯LEDn", "1号梯照明指示" => "输出"."2号梯照明指示", "1号梯风扇指示" => "输出"."2号梯风扇指示", "1号梯满载指示" => "输出"."2号梯满载指示", "1号梯故障指示" => "输出"."2号梯故障指示")
   END_RUNG
   // the same network as SCL:
   "2号梯指示灯"("1号梯光幕信号" := "输入"."2号梯光幕信号",   // "照明，风扇，数码管"
            "1号梯开门到位" := "输入"."2号梯开门到位",
            "1号梯当前载重量" := "中间变量2"."2号梯转换后载重量",
            当前楼层数 := "中间变量1"."2号梯当前楼层数",
            "1号梯检修信号" := "输入"."2号梯检修信号",
            开门继电器 := "输出"."2号梯开门继电器",
            关门继电器 := "输出"."2号梯关门继电器",
            关门到位 := "输入"."2号梯关门到位",
            转换后载重量 := "中间变量2"."2号梯转换后载重量",
            载重限额 := "中间变量1"."2号梯载重限额",
            上行接触器 := "输出"."2号梯上行接触器",
            下行接触器 := "输出"."2号梯下行接触器",
            正处于故障中 => "中间变量1"."2号梯正处于故障中",
            安全隐患 => "中间变量1"."2号梯存在安全隐患（光幕）",
            "1号梯LEDa" => "输出"."2号梯LEDa",
            "1号梯LEDb" => "输出"."2号梯LEDb",
            "1号梯LEDc" => "输出"."2号梯LEDc",
            "1号梯LEDd" => "输出"."2号梯LEDd",
            "1号梯LEDe" => "输出"."2号梯LEDe",
            "1号梯LEDf" => "输出"."2号梯LEDf",
            "1号梯LEDg" => "输出"."2号梯LEDg",
            "1号梯LEDh" => "输出"."2号梯LEDh",
            "1号梯LEDi" => "输出"."2号梯LEDi",
            "1号梯LEDj" => "输出"."2号梯LEDj",
            "1号梯LEDk" => "输出"."2号梯LEDk",
            "1号梯LEDl" => "输出"."2号梯LEDl",
            "1号梯LEDm" => "输出"."2号梯LEDm",
            "1号梯LEDn" => "输出"."2号梯LEDn",
            "1号梯照明指示" => "输出"."2号梯照明指示",
            "1号梯风扇指示" => "输出"."2号梯风扇指示",
            "1号梯满载指示" => "输出"."2号梯满载指示",
            "1号梯故障指示" => "输出"."2号梯故障指示");
END_REGION

REGION Network 3: 3号梯指示灯
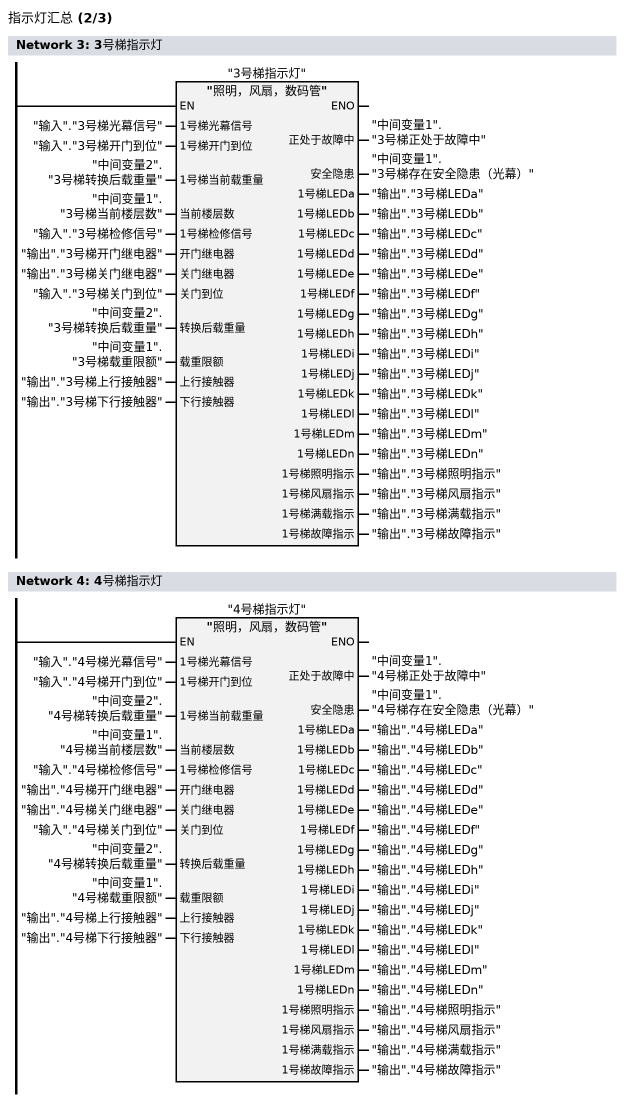
   RUNG wire#powerrail
      "3号梯指示灯"("1号梯光幕信号" := "输入"."3号梯光幕信号", "1号梯开门到位" := "输入"."3号梯开门到位", "1号梯当前载重量" := "中间变量2"."3号梯转换后载重量", 当前楼层数 := "中间变量1"."3号梯当前楼层数", "1号梯检修信号" := "输入"."3号梯检修信号", 开门继电器 := "输出"."3号梯开门继电器", 关门继电器 := "输出"."3号梯关门继电器", 关门到位 := "输入"."3号梯关门到位", 转换后载重量 := "中间变量2"."3号梯转换后载重量", 载重限额 := "中间变量1"."3号梯载重限额", 上行接触器 := "输出"."3号梯上行接触器", 下行接触器 := "输出"."3号梯下行接触器", 正处于故障中 => "中间变量1"."3号梯正处于故障中", 安全隐患 => "中间变量1"."3号梯存在安全隐患（光幕）", "1号梯LEDa" => "输出"."3号梯LEDa", "1号梯LEDb" => "输出"."3号梯LEDb", "1号梯LEDc" => "输出"."3号梯LEDc", "1号梯LEDd" => "输出"."3号梯LEDd", "1号梯LEDe" => "输出"."3号梯LEDe", "1号梯LEDf" => "输出"."3号梯LEDf", "1号梯LEDg" => "输出"."3号梯LEDg", "1号梯LEDh" => "输出"."3号梯LEDh", "1号梯LEDi" => "输出"."3号梯LEDi", "1号梯LEDj" => "输出"."3号梯LEDj", "1号梯LEDk" => "输出"."3号梯LEDk", "1号梯LEDl" => "输出"."3号梯LEDl", "1号梯LEDm" => "输出"."3号梯LEDm", "1号梯LEDn" => "输出"."3号梯LEDn", "1号梯照明指示" => "输出"."3号梯照明指示", "1号梯风扇指示" => "输出"."3号梯风扇指示", "1号梯满载指示" => "输出"."3号梯满载指示", "1号梯故障指示" => "输出"."3号梯故障指示")
   END_RUNG
   // the same network as SCL:
   "3号梯指示灯"("1号梯光幕信号" := "输入"."3号梯光幕信号",   // "照明，风扇，数码管"
            "1号梯开门到位" := "输入"."3号梯开门到位",
            "1号梯当前载重量" := "中间变量2"."3号梯转换后载重量",
            当前楼层数 := "中间变量1"."3号梯当前楼层数",
            "1号梯检修信号" := "输入"."3号梯检修信号",
            开门继电器 := "输出"."3号梯开门继电器",
            关门继电器 := "输出"."3号梯关门继电器",
            关门到位 := "输入"."3号梯关门到位",
            转换后载重量 := "中间变量2"."3号梯转换后载重量",
            载重限额 := "中间变量1"."3号梯载重限额",
            上行接触器 := "输出"."3号梯上行接触器",
            下行接触器 := "输出"."3号梯下行接触器",
            正处于故障中 => "中间变量1"."3号梯正处于故障中",
            安全隐患 => "中间变量1"."3号梯存在安全隐患（光幕）",
            "1号梯LEDa" => "输出"."3号梯LEDa",
            "1号梯LEDb" => "输出"."3号梯LEDb",
            "1号梯LEDc" => "输出"."3号梯LEDc",
            "1号梯LEDd" => "输出"."3号梯LEDd",
            "1号梯LEDe" => "输出"."3号梯LEDe",
            "1号梯LEDf" => "输出"."3号梯LEDf",
            "1号梯LEDg" => "输出"."3号梯LEDg",
            "1号梯LEDh" => "输出"."3号梯LEDh",
            "1号梯LEDi" => "输出"."3号梯LEDi",
            "1号梯LEDj" => "输出"."3号梯LEDj",
            "1号梯LEDk" => "输出"."3号梯LEDk",
            "1号梯LEDl" => "输出"."3号梯LEDl",
            "1号梯LEDm" => "输出"."3号梯LEDm",
            "1号梯LEDn" => "输出"."3号梯LEDn",
            "1号梯照明指示" => "输出"."3号梯照明指示",
            "1号梯风扇指示" => "输出"."3号梯风扇指示",
            "1号梯满载指示" => "输出"."3号梯满载指示",
            "1号梯故障指示" => "输出"."3号梯故障指示");
END_REGION

REGION Network 4: 4号梯指示灯
   RUNG wire#powerrail
      "4号梯指示灯"("1号梯光幕信号" := "输入"."4号梯光幕信号", "1号梯开门到位" := "输入"."4号梯开门到位", "1号梯当前载重量" := "中间变量2"."4号梯转换后载重量", 当前楼层数 := "中间变量1"."4号梯当前楼层数", "1号梯检修信号" := "输入"."4号梯检修信号", 开门继电器 := "输出"."4号梯开门继电器", 关门继电器 := "输出"."4号梯关门继电器", 关门到位 := "输入"."4号梯关门到位", 转换后载重量 := "中间变量2"."4号梯转换后载重量", 载重限额 := "中间变量1"."4号梯载重限额", 上行接触器 := "输出"."4号梯上行接触器", 下行接触器 := "输出"."4号梯下行接触器", 正处于故障中 => "中间变量1"."4号梯正处于故障中", 安全隐患 => "中间变量1"."4号梯存在安全隐患（光幕）", "1号梯LEDa" => "输出"."4号梯LEDa", "1号梯LEDb" => "输出"."4号梯LEDb", "1号梯LEDc" => "输出"."4号梯LEDc", "1号梯LEDd" => "输出"."4号梯LEDd", "1号梯LEDe" => "输出"."4号梯LEDe", "1号梯LEDf" => "输出"."4号梯LEDf", "1号梯LEDg" => "输出"."4号梯LEDg", "1号梯LEDh" => "输出"."4号梯LEDh", "1号梯LEDi" => "输出"."4号梯LEDi", "1号梯LEDj" => "输出"."4号梯LEDj", "1号梯LEDk" => "输出"."4号梯LEDk", "1号梯LEDl" => "输出"."4号梯LEDl", "1号梯LEDm" => "输出"."4号梯LEDm", "1号梯LEDn" => "输出"."4号梯LEDn", "1号梯照明指示" => "输出"."4号梯照明指示", "1号梯风扇指示" => "输出"."4号梯风扇指示", "1号梯满载指示" => "输出"."4号梯满载指示", "1号梯故障指示" => "输出"."4号梯故障指示")
   END_RUNG
   // the same network as SCL:
   "4号梯指示灯"("1号梯光幕信号" := "输入"."4号梯光幕信号",   // "照明，风扇，数码管"
            "1号梯开门到位" := "输入"."4号梯开门到位",
            "1号梯当前载重量" := "中间变量2"."4号梯转换后载重量",
            当前楼层数 := "中间变量1"."4号梯当前楼层数",
            "1号梯检修信号" := "输入"."4号梯检修信号",
            开门继电器 := "输出"."4号梯开门继电器",
            关门继电器 := "输出"."4号梯关门继电器",
            关门到位 := "输入"."4号梯关门到位",
            转换后载重量 := "中间变量2"."4号梯转换后载重量",
            载重限额 := "中间变量1"."4号梯载重限额",
            上行接触器 := "输出"."4号梯上行接触器",
            下行接触器 := "输出"."4号梯下行接触器",
            正处于故障中 => "中间变量1"."4号梯正处于故障中",
            安全隐患 => "中间变量1"."4号梯存在安全隐患（光幕）",
            "1号梯LEDa" => "输出"."4号梯LEDa",
            "1号梯LEDb" => "输出"."4号梯LEDb",
            "1号梯LEDc" => "输出"."4号梯LEDc",
            "1号梯LEDd" => "输出"."4号梯LEDd",
            "1号梯LEDe" => "输出"."4号梯LEDe",
            "1号梯LEDf" => "输出"."4号梯LEDf",
            "1号梯LEDg" => "输出"."4号梯LEDg",
            "1号梯LEDh" => "输出"."4号梯LEDh",
            "1号梯LEDi" => "输出"."4号梯LEDi",
            "1号梯LEDj" => "输出"."4号梯LEDj",
            "1号梯LEDk" => "输出"."4号梯LEDk",
            "1号梯LEDl" => "输出"."4号梯LEDl",
            "1号梯LEDm" => "输出"."4号梯LEDm",
            "1号梯LEDn" => "输出"."4号梯LEDn",
            "1号梯照明指示" => "输出"."4号梯照明指示",
            "1号梯风扇指示" => "输出"."4号梯风扇指示",
            "1号梯满载指示" => "输出"."4号梯满载指示",
            "1号梯故障指示" => "输出"."4号梯故障指示");
END_REGION

REGION Network 5: 5号梯指示灯
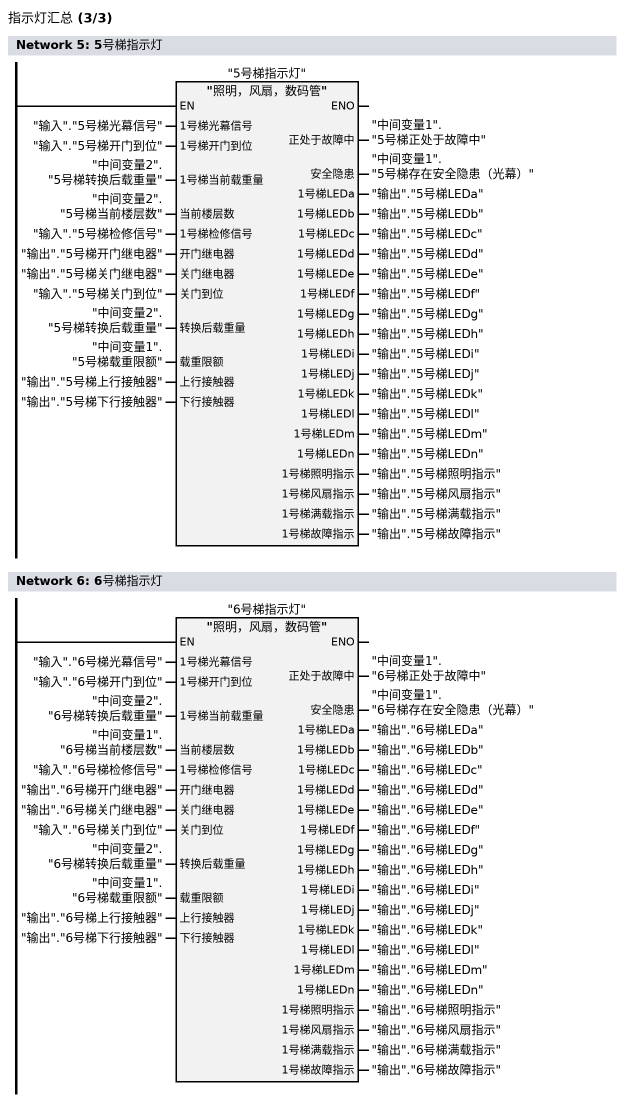
   RUNG wire#powerrail
      "5号梯指示灯"("1号梯光幕信号" := "输入"."5号梯光幕信号", "1号梯开门到位" := "输入"."5号梯开门到位", "1号梯当前载重量" := "中间变量2"."5号梯转换后载重量", 当前楼层数 := "中间变量2"."5号梯当前楼层数", "1号梯检修信号" := "输入"."5号梯检修信号", 开门继电器 := "输出"."5号梯开门继电器", 关门继电器 := "输出"."5号梯关门继电器", 关门到位 := "输入"."5号梯关门到位", 转换后载重量 := "中间变量2"."5号梯转换后载重量", 载重限额 := "中间变量1"."5号梯载重限额", 上行接触器 := "输出"."5号梯上行接触器", 下行接触器 := "输出"."5号梯下行接触器", 正处于故障中 => "中间变量1"."5号梯正处于故障中", 安全隐患 => "中间变量1"."5号梯存在安全隐患（光幕）", "1号梯LEDa" => "输出"."5号梯LEDa", "1号梯LEDb" => "输出"."5号梯LEDb", "1号梯LEDc" => "输出"."5号梯LEDc", "1号梯LEDd" => "输出"."5号梯LEDd", "1号梯LEDe" => "输出"."5号梯LEDe", "1号梯LEDf" => "输出"."5号梯LEDf", "1号梯LEDg" => "输出"."5号梯LEDg", "1号梯LEDh" => "输出"."5号梯LEDh", "1号梯LEDi" => "输出"."5号梯LEDi", "1号梯LEDj" => "输出"."5号梯LEDj", "1号梯LEDk" => "输出"."5号梯LEDk", "1号梯LEDl" => "输出"."5号梯LEDl", "1号梯LEDm" => "输出"."5号梯LEDm", "1号梯LEDn" => "输出"."5号梯LEDn", "1号梯照明指示" => "输出"."5号梯照明指示", "1号梯风扇指示" => "输出"."5号梯风扇指示", "1号梯满载指示" => "输出"."5号梯满载指示", "1号梯故障指示" => "输出"."5号梯故障指示")
   END_RUNG
   // the same network as SCL:
   "5号梯指示灯"("1号梯光幕信号" := "输入"."5号梯光幕信号",   // "照明，风扇，数码管"
            "1号梯开门到位" := "输入"."5号梯开门到位",
            "1号梯当前载重量" := "中间变量2"."5号梯转换后载重量",
            当前楼层数 := "中间变量2"."5号梯当前楼层数",
            "1号梯检修信号" := "输入"."5号梯检修信号",
            开门继电器 := "输出"."5号梯开门继电器",
            关门继电器 := "输出"."5号梯关门继电器",
            关门到位 := "输入"."5号梯关门到位",
            转换后载重量 := "中间变量2"."5号梯转换后载重量",
            载重限额 := "中间变量1"."5号梯载重限额",
            上行接触器 := "输出"."5号梯上行接触器",
            下行接触器 := "输出"."5号梯下行接触器",
            正处于故障中 => "中间变量1"."5号梯正处于故障中",
            安全隐患 => "中间变量1"."5号梯存在安全隐患（光幕）",
            "1号梯LEDa" => "输出"."5号梯LEDa",
            "1号梯LEDb" => "输出"."5号梯LEDb",
            "1号梯LEDc" => "输出"."5号梯LEDc",
            "1号梯LEDd" => "输出"."5号梯LEDd",
            "1号梯LEDe" => "输出"."5号梯LEDe",
            "1号梯LEDf" => "输出"."5号梯LEDf",
            "1号梯LEDg" => "输出"."5号梯LEDg",
            "1号梯LEDh" => "输出"."5号梯LEDh",
            "1号梯LEDi" => "输出"."5号梯LEDi",
            "1号梯LEDj" => "输出"."5号梯LEDj",
            "1号梯LEDk" => "输出"."5号梯LEDk",
            "1号梯LEDl" => "输出"."5号梯LEDl",
            "1号梯LEDm" => "输出"."5号梯LEDm",
            "1号梯LEDn" => "输出"."5号梯LEDn",
            "1号梯照明指示" => "输出"."5号梯照明指示",
            "1号梯风扇指示" => "输出"."5号梯风扇指示",
            "1号梯满载指示" => "输出"."5号梯满载指示",
            "1号梯故障指示" => "输出"."5号梯故障指示");
END_REGION

REGION Network 6: 6号梯指示灯
   RUNG wire#powerrail
      "6号梯指示灯"("1号梯光幕信号" := "输入"."6号梯光幕信号", "1号梯开门到位" := "输入"."6号梯开门到位", "1号梯当前载重量" := "中间变量2"."6号梯转换后载重量", 当前楼层数 := "中间变量1"."6号梯当前楼层数", "1号梯检修信号" := "输入"."6号梯检修信号", 开门继电器 := "输出"."6号梯开门继电器", 关门继电器 := "输出"."6号梯关门继电器", 关门到位 := "输入"."6号梯关门到位", 转换后载重量 := "中间变量2"."6号梯转换后载重量", 载重限额 := "中间变量1"."6号梯载重限额", 上行接触器 := "输出"."6号梯上行接触器", 下行接触器 := "输出"."6号梯下行接触器", 正处于故障中 => "中间变量1"."6号梯正处于故障中", 安全隐患 => "中间变量1"."6号梯存在安全隐患（光幕）", "1号梯LEDa" => "输出"."6号梯LEDa", "1号梯LEDb" => "输出"."6号梯LEDb", "1号梯LEDc" => "输出"."6号梯LEDc", "1号梯LEDd" => "输出"."6号梯LEDd", "1号梯LEDe" => "输出"."6号梯LEDe", "1号梯LEDf" => "输出"."6号梯LEDf", "1号梯LEDg" => "输出"."6号梯LEDg", "1号梯LEDh" => "输出"."6号梯LEDh", "1号梯LEDi" => "输出"."6号梯LEDi", "1号梯LEDj" => "输出"."6号梯LEDj", "1号梯LEDk" => "输出"."6号梯LEDk", "1号梯LEDl" => "输出"."6号梯LEDl", "1号梯LEDm" => "输出"."6号梯LEDm", "1号梯LEDn" => "输出"."6号梯LEDn", "1号梯照明指示" => "输出"."6号梯照明指示", "1号梯风扇指示" => "输出"."6号梯风扇指示", "1号梯满载指示" => "输出"."6号梯满载指示", "1号梯故障指示" => "输出"."6号梯故障指示")
   END_RUNG
   // the same network as SCL:
   "6号梯指示灯"("1号梯光幕信号" := "输入"."6号梯光幕信号",   // "照明，风扇，数码管"
            "1号梯开门到位" := "输入"."6号梯开门到位",
            "1号梯当前载重量" := "中间变量2"."6号梯转换后载重量",
            当前楼层数 := "中间变量1"."6号梯当前楼层数",
            "1号梯检修信号" := "输入"."6号梯检修信号",
            开门继电器 := "输出"."6号梯开门继电器",
            关门继电器 := "输出"."6号梯关门继电器",
            关门到位 := "输入"."6号梯关门到位",
            转换后载重量 := "中间变量2"."6号梯转换后载重量",
            载重限额 := "中间变量1"."6号梯载重限额",
            上行接触器 := "输出"."6号梯上行接触器",
            下行接触器 := "输出"."6号梯下行接触器",
            正处于故障中 => "中间变量1"."6号梯正处于故障中",
            安全隐患 => "中间变量1"."6号梯存在安全隐患（光幕）",
            "1号梯LEDa" => "输出"."6号梯LEDa",
            "1号梯LEDb" => "输出"."6号梯LEDb",
            "1号梯LEDc" => "输出"."6号梯LEDc",
            "1号梯LEDd" => "输出"."6号梯LEDd",
            "1号梯LEDe" => "输出"."6号梯LEDe",
            "1号梯LEDf" => "输出"."6号梯LEDf",
            "1号梯LEDg" => "输出"."6号梯LEDg",
            "1号梯LEDh" => "输出"."6号梯LEDh",
            "1号梯LEDi" => "输出"."6号梯LEDi",
            "1号梯LEDj" => "输出"."6号梯LEDj",
            "1号梯LEDk" => "输出"."6号梯LEDk",
            "1号梯LEDl" => "输出"."6号梯LEDl",
            "1号梯LEDm" => "输出"."6号梯LEDm",
            "1号梯LEDn" => "输出"."6号梯LEDn",
            "1号梯照明指示" => "输出"."6号梯照明指示",
            "1号梯风扇指示" => "输出"."6号梯风扇指示",
            "1号梯满载指示" => "输出"."6号梯满载指示",
            "1号梯故障指示" => "输出"."6号梯故障指示");
END_REGION
END_FUNCTION

FUNCTION "电梯目标判断" : Void   // FC12, LAD
{ S7_Optimized_Access := 'TRUE' }
VERSION : 0.1
BEGIN

REGION Network 2
